        IF NOT _done THEN
            _to_A._sut_A.Invoke();
            _to_A._sut_B.Invoke();
            _to_A();

            IF _to_A._sut_A.Done AND NOT _retBool THEN
                _to_A._sut_A.Abort();
                _to_A._sut_B.Abort();
                _retBool := true;
            END_IF

            _done := _to_A._sut_A.Done AND _to_A._sut_B.Done;
        END_IF

        IF _done THEN
            _to_A._sut_A.ReadOutState();
            _to_A._sut_B.ReadOutState();
            ProbeDoneWhen(_done);
        END_IF
    {endregion}
    {region "T310_TaskError"}
    eTcoTaskTests.TaskError:
        IF NOT _arranged THEN
            IF _plcCycleCounter = 1 THEN
                _to_A.CounterValue_A := _inUint;
                RETURN;
            END_IF

            IF _plcCycleCounter = 2 THEN
                _to_A._sut_A.Invoke();
                RETURN;
            END_IF

            IF _plcCycleCounter > 2 AND _plcCycleCounter <= 5 THEN
                _to_A._sut_A();
                RETURN;
            END_IF

            IF _plcCycleCounter = 6 THEN
                _to_A._sut_A();
                _to_A._sut_A.ReadOutState();
                _arranged := TRUE;
                RETURN;
            END_IF
        END_IF

        IF NOT _done THEN
            IF _plcCycleCounter = 7 THEN
                _to_A.CounterValue_A := _to_A.CounterValue_A + 5;
                _to_A._sut_A();
                _to_A._sut_A.ReadOutState();
            END_IF

            IF _plcCycleCounter > 7 AND _plcCycleCounter <= 7 + _inUint THEN
                _to_A._sut_A();
                _to_A._sut_A.ReadOutState();
            END_IF

            _done := _plcCycleCounter >= 7 + _inUint;
            ProbeDoneWhen(_done);
        END_IF
    {endregion}
    {region "T311_TaskInvokeAfterErrorNoRestoreNoEmptyCycles"}
    eTcoTaskTests.TaskInvokeAfterErrorNoRestoreNoEmptyCycles:
        IF NOT _arranged THEN
            _to_A._sut_A.Invoke();
            _arranged := TRUE;
            RETURN;
        END_IF

        IF NOT _done THEN
            _to_A._sut_A();
            _to_A._sut_A.ReadOutState();
            ProbeDoneWhen(_plcCycleCounter >= 1 + _inUint);
        END_IF
    {endregion}
    {region "T312_TaskInvokeAfterErrorNoRestoreOneEmptyCycle"}
    eTcoTaskTests.TaskInvokeAfterErrorNoRestoreOneEmptyCycle:
        IF NOT _arranged THEN
            IF _plcCycleCounter = 1 THEN
                RETURN;
            END_IF

            IF _plcCycleCounter = 2 THEN
                _to_A._sut_A.Invoke();
                RETURN;
            END_IF
        END_IF

        IF NOT _done THEN
            _to_A._sut_A();
            _to_A._sut_A.ReadOutState();
            _done := _plcCycleCounter >= 2 + _inUint;
            ProbeDoneWhen(_done);
        END_IF
    {endregion}
    {region "T313_TaskInvokeAfterErrorWithRestore"}
    eTcoTaskTests.TaskInvokeAfterErrorWithRestore:
        _to_A._sut_A.Restore();
        _to_A._sut_A.Invoke();
        _to_A._sut_A();
        _to_A._sut_A.ReadOutState();
        _done := TRUE;
        ProbeDoneWhen(_done);
    {endregion}
    {region "T314_TaskAbortDuringExecution"}
    eTcoTaskTests.TaskAbortDuringExecution:
        IF _plcCycleCounter = 1 THEN
            _to_A._sut_A.Restore();
            RETURN;
        END_IF

        IF _plcCycleCounter = 2 THEN
            _to_A._sut_A.Invoke();
            _to_A._sut_A();
            _to_A._sut_A.ReadOutState();
            RETURN;
        END_IF

        IF _plcCycleCounter = 3 THEN
            _to_A._sut_A.Abort();
            _to_A._sut_A();
            _to_A._sut_A.ReadOutState();
            _done := TRUE;
            ProbeDoneWhen(_done);
        END_IF
    {endregion}
    {region "T315_TaskMessage"}
    eTcoTaskTests.TaskMessage:
        _to_A._sut_A.PostMessage(Message := _inString);
        _retString := _to_A._sut_A.GetMessage();
        _done := TRUE;
        ProbeDoneWhen(_done);
    {endregion}
    {region "T316_IdentitiesTest"}
    eTcoTaskTests.IdentitiesTest:
        _runElapsedTimer := TRUE;
        _elapsedTimeETA := UINT_TO_TIME(_inUint);
        _to_A._sut_A.ReadOutIdentities();
        _to_A.ReadOutIdentities();
        ReadOutCycleCounters();
        _done := _elapsedTimeTimer.Q;
        ProbeDoneWhen(_done);
    {endregion}
    {region "T317_CheckAutoRestoreProperties"}
    eTcoTaskTests.CheckAutoRestoreProperties:
        _to_A._tSt_A.ReadOutAutoRestoreProperties();
        _to_A._tSt_B.ReadOutAutoRestoreProperties();
        _to_A._tSt_A._tTt_A.ReadOutAutoRestoreProperties();
        _to_A._tSt_A._tTt_B.ReadOutAutoRestoreProperties();
        _to_A._tSt_B._tTt_A.ReadOutAutoRestoreProperties();
        _to_A._tSt_B._tTt_B.ReadOutAutoRestoreProperties();
        _done := TRUE;
        ProbeDoneWhen(_done);
    {endregion}
    {region "T318_AutoRestoreOnStateChange"}
    eTcoTaskTests.AutoRestoreOnStateChange:
        IF _plcCycleCounter = 1 THEN
            _to_A._tSt_A.ReadOutAutoRestoreProperties();
            _to_A._tSt_B.ReadOutAutoRestoreProperties();
            _to_A._tSt_A._tTt_A.ReadOutAutoRestoreProperties();
            _to_A._tSt_A._tTt_B.ReadOutAutoRestoreProperties();
            _to_A._tSt_B._tTt_A.ReadOutAutoRestoreProperties();
            _to_A._tSt_B._tTt_B.ReadOutAutoRestoreProperties();
            _to_A._tSt_A._tTt_A.ReadOutState();
            _to_A._tSt_B._tTt_B.ReadOutState();
        END_IF

        IF _plcCycleCounter = 2 THEN
            _to_A._tSt_A._tTt_A.Restore();
            _to_A._tSt_B._tTt_B.Restore();
            _to_A._tSt_A._tTt_A.ReadOutState();
            _to_A._tSt_B._tTt_B.ReadOutState();
        END_IF

        IF _plcCycleCounter = 3 THEN
            _to_A._tSt_A._tTt_A.Invoke();
            _to_A._tSt_B._tTt_B.Invoke();
            _to_A._tSt_A._tTt_A();
            _to_A._tSt_B._tTt_B();
            _to_A._tSt_A._tTt_A.ReadOutState();
            _to_A._tSt_B._tTt_B.ReadOutState();
        END_IF

        IF _plcCycleCounter = 4 THEN
            _to_A._tSt_A._tTt_A.Invoke();
            _to_A._tSt_A._tTt_A();
            _to_A._tSt_B._tTt_B();
            _to_A._tSt_A._tTt_A.ReadOutState();
            _to_A._tSt_B._tTt_B.ReadOutState();
        END_IF

        IF _plcCycleCounter = 5 THEN
            _to_A._tSt_A.ChangeState(_to_A._tSt_A._myState);
            _to_A._tSt_B.ChangeState(_to_A._tSt_B._myState);
            _to_A._tSt_A._tTt_A();
            _to_A._tSt_B._tTt_B();
            _to_A._tSt_A._tTt_A.ReadOutState();
            _to_A._tSt_B._tTt_B.ReadOutState();
        END_IF

        _done := _plcCycleCounter = 5;
        ProbeDoneWhen(_done);
    {endregion}
    {region "T320_InvokeDisabledTask"}
    eTcoTaskTests.InvokeDisabledTask:
        IF _plcCycleCounter = 1 THEN
            _to_A._sut_A.Restore();
            _to_A._sut_A.Disable();
            RETURN;
        END_IF

        IF NOT _done THEN
            _to_A._sut_A.Invoke();
            _to_A._sut_A();
            _to_A._sut_A.ReadOutState();
            _done := _plcCycleCounter >= 1 + _inUint;
            ProbeDoneWhen(_done);
        END_IF
    {endregion}
    {region "T321_DisableExecutingTask"}
    eTcoTaskTests.DisableExecutingTask:
        IF _plcCycleCounter = 1 THEN
            _to_A._sut_A.Enable();
            _to_A._sut_A.Invoke();
            _to_A._sut_A();
            _to_A._sut_A.ReadOutState();
            RETURN;
        END_IF

        IF _plcCycleCounter = 2 THEN
            _to_A._sut_A.Disable();
            _to_A._sut_A();
            _to_A._sut_A.ReadOutState();
            RETURN;
        END_IF

        IF _plcCycleCounter = 3 THEN
            _to_A._sut_A.Restore();
            _to_A._sut_A.Enable();
            _to_A._sut_A();
            _to_A._sut_A.ReadOutState();
            RETURN;
        END_IF

        IF _plcCycleCounter = 4 THEN
            _to_A._sut_A.Invoke();
            _to_A._sut_A();
            _to_A._sut_A.ReadOutState();
            RETURN;
        END_IF

        IF _plcCycleCounter = 5 THEN
            _to_A._sut_A.Restore();
            _to_A._sut_A();
            _to_A._sut_A.ReadOutState();
            _done := TRUE;
            ProbeDoneWhen(_done);
        END_IF
    {endregion}
    {region "T322_InvokeTaskThenDisable"}
    eTcoTaskTests.InvokeTaskThenDisable:
        _to_A._sut_A.Invoke();
        _to_A._sut_A.Disable();
        _to_A._sut_A();
        _to_A._sut_A.ReadOutState();
        _done := TRUE;
        ProbeDoneWhen(_done);
    {endregion}
    {region "T323_DisableTaskInErrorStateEnableAndTriggerAgain"}
    eTcoTaskTests.DisableTaskInErrorStateEnableAndTriggerAgain:
        IF _plcCycleCounter = 1 THEN
            _to_A._sut_A.Enable();
            _to_A._sut_A.Invoke();
            _to_A._sut_A();
            _to_A._sut_A.ReadOutState();
            RETURN;
        END_IF

        IF _plcCycleCounter = 2 THEN
            _to_A.CounterValue_A := _to_A.CounterValue_A + 5;
            _to_A._sut_A();
            _to_A._sut_A.ReadOutState();
            RETURN;
        END_IF

        IF _plcCycleCounter = 3 THEN
            _to_A._sut_A.Disable();
            _to_A._sut_A();
            _to_A._sut_A.ReadOutState();
            RETURN;
        END_IF

        IF _plcCycleCounter = 4 THEN
            _to_A._sut_A.Invoke();
            _to_A._sut_A();
            _to_A._sut_A.ReadOutState();
            RETURN;
        END_IF

        IF _plcCycleCounter = 5 THEN
            _to_A._sut_A.Restore();
            _to_A._sut_A.Invoke();
            _to_A._sut_A();
            _to_A._sut_A.ReadOutState();
            _done := TRUE;
            ProbeDoneWhen(_done);
        END_IF
    {endregion}
    {region "T330_ElapsedTypeMeasurement"}
    eTcoTaskTests.ElapsedTypeMeasurement:
        IF _plcCycleCounter = 1 THEN
            _to_A._sut_A.Restore();
            _to_A._sut_A.Enable();
            _to_A._sut_A.Invoke();
            RETURN;
        END_IF

        IF (_to_A._sut_A.Execute()) THEN
            _runElapsedTimer := TRUE;

            IF (_elapsedTimeTimer.Q) THEN
                _to_A._sut_A.DoneWhen(_elapsedTimeTimer.Q);
            END_IF;
        END_IF

        _done := _to_A._sut_A.Done;
        ProbeDoneWhen(_done);
        _elapsedTime := _to_A._sut_A.ElapsedTime;
    {endregion}
    {region "T340_TaskExecutingWithDoneAndErrorStatement"}
    eTcoTaskTests.TaskExecutingWithDoneAndErrorStatement:
        IF _plcCycleCounter = 1 THEN
            _to_A._sut_A.Restore();
            _to_A._sut_A.Enable();
            _to_A._sut_A.Invoke();
            _to_A._sut_A();
            _to_A._sut_A.ReadOutState();
            RETURN;
        END_IF

        _to_A._sut_A();
        _to_A._sut_A.DoneWhen(TRUE);
        _to_A._sut_A.ThrowWhen(TRUE);
        _to_A._sut_A.ReadOutState();
        _done := _to_A._sut_A.Done;
        ProbeDoneWhen(_done);
    {endregion}
    {region "T341_TaskExecutingWithErrorAndDoneStatement"}
    eTcoTaskTests.TaskExecutingWithErrorAndDoneStatement:
        IF _plcCycleCounter = 1 THEN
            _to_A._sut_A.Restore();
            _to_A._sut_A.Enable();
            _to_A._sut_A.Invoke();
            _to_A._sut_A();
            _to_A._sut_A.ReadOutState();
            RETURN;
        END_IF

        _to_A._sut_A();
        _to_A._sut_A.ThrowWhen(TRUE);
        _to_A._sut_A.DoneWhen(TRUE);
        _to_A._sut_A.ReadOutState();
        _done := _to_A._sut_A.Done;
        ProbeDoneWhen(_done);			 
{endregion}
	 eTcoTaskTests.TaskExecuteMethodNotCalled:
	 	_to_A._sut_A.Invoke().Done;
	eTcoTaskTests.TaskExecuteMethodCalled :
		_to_A._sut_A.Invoke().Done;
		_to_A._sut_A.Execute();
END_CASE
END_METHOD

METHOD INTERNAL ReadOutCycleCounters
_startCycles		:=		THIS^.StartCycleCount;
_endCycles			:=		THIS^.EndCycleCount;

_myIdentity			:= 		THIS^.Identity;
END_METHOD

END_FUNCTION_BLOCK

// ---- Tests/TcoTask/PlcExecuted/TcoTaskPlcTestObject.TcPOU
FUNCTION_BLOCK TcoTaskPlcTestObject EXTENDS TcoCore.TcoObject
VAR
	_myIdentity				:	ULINT;
	_myContextIdentity		:	ULINT;
	_myContextStartCount 	:	ULINT;
	_myContextEndCount		:	ULINT;
	_myParentIdentity		:	ULINT;
    _sut_A : TcoTaskPlcTest(THIS^);
    _sut_B : TcoTaskPlcTest(THIS^);
	_tSt_A:TcoTaskPlcTestState(THIS^, eRestoreMode.AutoRestoreMembers);
	_tSt_B:TcoTaskPlcTestState(THIS^, eRestoreMode.None);
END_VAR

_sut_A();
_sut_B();

PROPERTY CounterValue_A : ULINT
GET
CounterValue_A := _sut_A.CounterValue;
END_GET
SET
_sut_A.CounterValue := CounterValue_A;
END_SET
END_PROPERTY

PROPERTY CounterValue_B : ULINT
GET
CounterValue_B := _sut_B.CounterValue;
END_GET
SET
_sut_B.CounterValue := CounterValue_B;
END_SET
END_PROPERTY

{attribute 'TcRpcEnable'}
METHOD INTERNAL ReadOutIdentities
_myIdentity			:=	THIS^.Identity;

_myContextIdentity	:=	THIS^.Context.Identity;
		
_myContextStartCount :=	THIS^.Context.StartCycleCount;

_myContextEndCount	:=	THIS^.Context.EndCycleCount;

_myParentIdentity	:=	THIS^.Parent.Identity;
END_METHOD

END_FUNCTION_BLOCK

// ---- Tests/TcoTask/PlcExecuted/TcoTaskPlcTest.TcPOU
FUNCTION_BLOCK TcoTaskPlcTest EXTENDS TcoCore.TcoTask
VAR
    _isBusy : BOOL;
    _isError : BOOL;
    _isDone : BOOL;
    _isReady : BOOL;
    _isInvokeRequestTrue : BOOL;
    _counterSetValue : ULINT;
    _counterValue : ULINT;
    _invokeCounter : ULINT;
    _executeCounter : ULINT;
    _doneCounter : ULINT;
    _invokeRisingEdgeCounter : ULINT;
    _executeRisingEdgeCounter : ULINT;
    _doneRisingEdgeCounter : ULINT;
    _previousState : eTaskState;
    _counterValuePV : ULINT;
    _myIdentity : ULINT;
    _myContextIdentity : ULINT;
    _myContextStartCount : ULINT;
    _myContextEndCount : ULINT;
    _myParentIdentity : ULINT;
    _autoRestoreByMyParentEnabled : BOOL;
    _onErrorCounter : ULINT;
    _whileErrorCounter : ULINT;
    _onStartCounter : ULINT;
END_VAR

IF(THIS^._taskState = eTaskState.Requested) THEN
	_invokeCounter := _invokeCounter + 1; 
END_IF;

IF(THIS^._taskState = eTaskState.Requested AND _PreviousState <> eTaskState.Requested) THEN
	_counterValue	:=	_counterSetValue;
	_counterValuePV := _counterValue;
	_invokeRisingEdgeCounter := _invokeRisingEdgeCounter + 1;
END_IF

IF(THIS^._taskState = eTaskState.Busy AND _previousState <> eTaskState.Busy) THEN
	_executeRisingEdgeCounter := _executeRisingEdgeCounter + 1;
END_IF

_previousState	:=	THIS^._taskState;

IF(Execute()) THEN
	_executeCounter := _executeCounter + 1;	
	_counterValue := _counterValue - 1;
	DoneWhen(_counterValue <= 0);			
	ThrowWhen(ABS(_counterValuePV -_counterValue) > 1);
	_CounterValuePV := _counterValue;
END_IF

IF(THIS^._taskState = eTaskState.Done) THEN
	_doneCounter := _doneCounter + 1; 
END_IF;

IF(THIS^._taskState = eTaskState.Done AND _previousState <> eTaskState.Done) THEN
	_doneRisingEdgeCounter := _doneRisingEdgeCounter + 1; 
END_IF

PROPERTY CounterValue : ULINT
GET
CounterValue := _counterValue;
END_GET
SET
_counterValue := CounterValue;
END_SET
END_PROPERTY

METHOD INTERNAL Disable
THIS^.Enabled := FALSE;
END_METHOD

METHOD INTERNAL Enable
THIS^.Enabled := TRUE;
END_METHOD

METHOD INTERNAL GetMessage : STRING
GetMessage := SUPER^._messenger._mime.Text;
END_METHOD

METHOD PROTECTED OnError
_onErrorCounter := _onErrorCounter +1;
END_METHOD

METHOD PROTECTED OnStart
_onStartCounter := _onStartCounter +1;
END_METHOD

METHOD INTERNAL PostMessage
VAR_INPUT
	Message	:	STRING;
END_VAR
THIS^.Messenger.Post(Message ,eMessageCategory.Error);
END_METHOD

{attribute 'TcRpcEnable'}
METHOD INTERNAL ReadOutAutoRestoreProperties
_autoRestoreByMyParentEnabled	:= THIS^.AutoRestorable;
END_METHOD

{attribute 'TcRpcEnable'}
METHOD INTERNAL ReadOutIdentities
_myIdentity			:=	THIS^.Identity;
 
_myContextIdentity	:=	THIS^.Context.Identity;
		
_myContextStartCount :=	THIS^.Context.StartCycleCount;
 
_myContextEndCount	:=	THIS^.Context.EndCycleCount;
 
_myParentIdentity	:=	THIS^.Parent.Identity;
END_METHOD

{attribute 'TcRpcEnable'}
METHOD INTERNAL ReadOutState
_isBusy					:=	THIS^.Busy;	
_isError				:=	THIS^.Error;	
_isDone					:=	THIS^.Done;	
_isReady				:=	THIS^.Ready;
_isInvokeRequestTrue 	:=	THIS^._invokeRequest;
END_METHOD

{attribute 'TcRpcEnable'}
METHOD INTERNAL SetInvokeRequest
THIS^._invokeRequest := TRUE;
END_METHOD

{attribute 'TcRpcEnable'}
METHOD INTERNAL SetPreviousStateToReady
THIS^._previousState := eTaskState.Ready;
END_METHOD

(*~
	<docu>
		<summary>
			Executes until task is in ```Error``` state .
		</summary>			
	</docu>	
~*)
METHOD PROTECTED WhileError
_whileErrorCounter := _whileErrorCounter + 1;
END_METHOD

END_FUNCTION_BLOCK

// ---- Tests/TcoTask/PlcExecuted/TcoTaskPlcTestState.TcPOU
FUNCTION_BLOCK TcoTaskPlcTestState EXTENDS TcoState
VAR
    _myIdentity : ULINT;
    _myContextIdentity : ULINT;
    _myContextStartCount : ULINT;
    _myContextEndCount : ULINT;
    _myParentIdentity : ULINT;
    _myState : INT;
    _tTt_A : TcoTaskPlcTest(THIS^);
    _tTt_B : TcoTaskPlcTest(THIS^);
    _onStateChangeCounter : INT;
    _autoRestoreToMyChildsEnabled : BOOL;
    _autoRestoreByMyParentEnabled : BOOL;
END_VAR

METHOD PROTECTED OnStateChange 
VAR_INPUT
	PreviousState	: INT;
	NewState 		: INT;
END_VAR
VAR
	message	:	STRING;
END_VAR
_onStateChangeCounter	:=	_onStateChangeCounter + 1;

message := CONCAT('My state has been change from ', INT_TO_STRING(PreviousState));
message := CONCAT(message, ' to the new state ');
message := CONCAT(message, INT_TO_STRING(NewState));
message := CONCAT(message, '.');

THIS^.Messenger.Post(message,eMessageCategory.Debug);

SUPER^.OnStateChange(PreviousState,NewState);
END_METHOD

{attribute 'TcRpcEnable'}
METHOD INTERNAL ReadOutAutoRestoreProperties
_autoRestoreToMyChildsEnabled	:= THIS^.IsAutoRestoreEnabled;
_autoRestoreByMyParentEnabled	:= THIS^.AutoRestorable;
END_METHOD

{attribute 'TcRpcEnable'}
METHOD INTERNAL ReadOutIdentities
_myIdentity			:=	THIS^.Identity;

_myContextIdentity	:=	THIS^.Context.Identity;

_myParentIdentity	:=	THIS^.Parent.Identity;
		
_myContextStartCount :=	THIS^.Context.StartCycleCount;

_myContextEndCount	:=	THIS^.Context.EndCycleCount;
END_METHOD

{attribute 'TcRpcEnable'}
METHOD INTERNAL ReadOutState
_myState			:=	THIS^.State;

THIS^._tTt_A.ReadOutState();
THIS^._tTt_B.ReadOutState();
END_METHOD

{attribute 'TcRpcEnable'}
METHOD INTERNAL TriggerChangeState
VAR_INPUT
	NewState : INT;
END_VAR
THIS^.ChangeState(NewState);
END_METHOD

{attribute 'TcRpcEnable'}
METHOD INTERNAL TriggerChangeStateWithObjectRestore
VAR_INPUT
	NewState : INT;
END_VAR
THIS^.ChangeState(NewState).RestoreObject(THIS^._tTt_A).RestoreObject(THIS^._tTt_B);
END_METHOD

{attribute 'TcRpcEnable'}
METHOD INTERNAL TriggerRestore
THIS^.Restore();
END_METHOD

{attribute 'TcRpcEnable'}
METHOD INTERNAL TriggerTaskInvoke
THIS^._tTt_A.Invoke();

THIS^._tTt_B.Invoke();
END_METHOD

END_FUNCTION_BLOCK

// ---- Tests/TcoToggleTask/TcoToggleTaskTestContext.TcPOU
FUNCTION_BLOCK TcoToggleTaskTestContext EXTENDS TcoCore._internals_TcoContext
VAR
    _sut 		:	TcoToggleTaskTests(THIS^, TRUE);
	_bool		:	BOOL;
	_string		:	STRING;
	_done		:	BOOL;
END_VAR

METHOD PROTECTED Main
CASE _testId OF
	eTcoToggleTaskTests.Reinit:
		_sut.FB_init(TRUE, FALSE, THIS^,_bool);
		_done := TRUE;
		
	eTcoToggleTaskTests.CleanUp:
		IF NOT _done THEN
			_sut._messenger.Clear();
			_done := TRUE;
		END_IF
		
	eTcoToggleTaskTests.Message:
		IF NOT _done THEN
			_sut.Messenger.Error(_string);
			_done := TRUE;
		END_IF
		
	eTcoToggleTaskTests.TriggerToggleWhileRunNotCalled:
		IF NOT _done THEN
			_sut._messenger.Clear();
			_sut.Toggle();
			_done := TRUE;	
		END_IF

	eTcoToggleTaskTests.TriggerToggleWhileDisabled:
		IF NOT _done THEN
			_sut.Run();
			_sut._messenger.Clear();
			_sut.Enabled := FALSE;
			_sut.Toggle();
			_done := TRUE;	
		END_IF

	eTcoToggleTaskTests.TriggerToggleWhileEnabled:
		IF NOT _done THEN
			_sut.Run();
			_sut._messenger.Clear();
			_sut.Enabled := TRUE;
			_sut.Toggle();
			_done := TRUE;	
		END_IF

	eTcoToggleTaskTests.TriggerOnWhileRunNotCalled:
		IF NOT _done THEN
			_sut._messenger.Clear();
			_sut.On();
			_done := TRUE;	
		END_IF

	eTcoToggleTaskTests.TriggerOnWhileDisabled:
		IF NOT _done THEN
			_sut.Run();
			_sut._messenger.Clear();
			_sut.Enabled := FALSE;
			_sut.On();
			_done := TRUE;	
		END_IF

	eTcoToggleTaskTests.TriggerOnWhileEnabled:
		IF NOT _done THEN
			_sut.Run();
			_sut._messenger.Clear();
			_sut.Enabled := TRUE;
			_sut.On();
			_done := TRUE;	
		END_IF

	eTcoToggleTaskTests.TriggerOffWhileRunNotCalled:
		IF NOT _done THEN
			_sut._messenger.Clear();
			_sut.Toggle();
			_done := TRUE;	
		END_IF

	eTcoToggleTaskTests.TriggerOffWhileDisabled:
		IF NOT _done THEN
			_sut.Run();
			_sut._messenger.Clear();
			_sut.Enabled := FALSE;
			_sut.Off();
			_done := TRUE;	
		END_IF

	eTcoToggleTaskTests.TriggerOffWhileEnabled:
		IF NOT _done THEN
			_sut.Run();
			_sut._messenger.Clear();
			_sut.Enabled := TRUE;
			_sut.Off();
			_done := TRUE;	
		END_IF

		
END_CASE
END_METHOD

END_FUNCTION_BLOCK

// ---- Tests/TcoToggleTask/TcoToggleTaskTests.TcPOU
FUNCTION_BLOCK TcoToggleTaskTests EXTENDS TcoCore.TcoToggleTask
VAR
	_isOn							:	BOOL;	
	_isOff							:	BOOL;	
	_isEnabled						:	BOOL;	
	_isToggleRequestTrue			:	BOOL;		
	_counterValue					:	ULINT;
	_counterValuePV					:	ULINT;
	_toggleCounter					:	ULINT;
	_runCounter						:	ULINT;
	_onFtrigCounter					:	ULINT;	
	_onRtrigCounter					:	ULINT;	
	_onCounter						:	ULINT;
	_offCounter						:	ULINT;
	_onStateChangeCounter			:	ULINT;
	_taskOnCounter					:	ULINT;
	_taskOffCounter					:	ULINT;
	_stateChangedCounter			:	ULINT;

	_previousState					:	BOOL;
	_myIdentity						:	ULINT;
	_myContextIdentity				:	ULINT;
	_myContextStartCount 			:	ULINT;
	_myContextEndCount				:	ULINT;	
	_myParentIdentity				:	ULINT;
END_VAR

ExecutionBody();

METHOD INTERNAL Disable
THIS^.Enabled := FALSE;
END_METHOD

METHOD INTERNAL Enable
THIS^.Enabled := TRUE;
END_METHOD

{attribute 'TcRpcEnable'}
METHOD INTERNAL ExecutionBody
Run();

_runCounter := _runCounter + 1;	

IF _previousState <> THIS^.State THEN
	_stateChangedCounter := _stateChangedCounter + 1;
END_IF; 
_previousState	:=	THIS^.State;
END_METHOD

{attribute 'TcRpcEnable'}
METHOD INTERNAL GetMessage : STRING
GetMessage := SUPER^._messenger._mime.Text;
END_METHOD

METHOD PROTECTED Main
VAR
	
END_VAR
END_METHOD

(*~
	<docu>
		<summary>
			Executes when toggle task changes its state from '''TRUE''' to '''FALSE'''.
		</summary>			
	</docu>	
~*)
METHOD PROTECTED OnFtrig
_onFtrigCounter := _onFtrigCounter + 1;
END_METHOD

(*~
	<docu>
		<summary>
			Executes when toggle task changes its state from '''FALSE''' to '''TRUE'''.
		</summary>			
	</docu>	
~*)
METHOD PROTECTED OnRtrig
_onRtrigCounter := _onRtrigCounter + 1;
END_METHOD

(*~
	<docu>
		<summary>
			Executes when toggle task changes its state .
		</summary>			
	</docu>	
~*)
METHOD PROTECTED OnStateChange
_onStateChangeCounter := _onStateChangeCounter + 1;
END_METHOD

{attribute 'TcRpcEnable'}
METHOD INTERNAL PostMessage
VAR_INPUT
	Message	:	STRING;
END_VAR
THIS^.Messenger.Post(Message ,eMessageCategory.Error);
END_METHOD

{attribute 'TcRpcEnable'}
METHOD INTERNAL ReadOutIdentities
_myIdentity			:=	THIS^.Identity;
 
_myContextIdentity	:=	THIS^.Context.Identity;
		
_myContextStartCount :=	THIS^.Context.StartCycleCount;
 
_myContextEndCount	:=	THIS^.Context.EndCycleCount;
 
_myParentIdentity	:=	THIS^.Parent.Identity;
END_METHOD

{attribute 'TcRpcEnable'}
METHOD INTERNAL ReadOutState
_isOn				    :=	THIS^.IsOn;	
_isOff				   	:=	THIS^.IsOff;	
_isEnabled				:=	THIS^.Enabled;
_isToggleRequestTrue	:=	THIS^._toggleRequest;
END_METHOD

{attribute 'TcRpcEnable'}
METHOD INTERNAL SetPreviousState
VAR_INPUT
	inValue : BOOL;
END_VAR
THIS^._previousState := inValue;
END_METHOD

{attribute 'TcRpcEnable'}
METHOD INTERNAL SetState
VAR_INPUT
	inState	:	BOOL;
END_VAR
THIS^._state := inState;
END_METHOD

{attribute 'TcRpcEnable'}
METHOD INTERNAL SetToggleRequest
THIS^._toggleRequest := TRUE;
END_METHOD

(*~
	<docu>
		<summary>
			Executes when toggle task is in ```Off``` state .
		</summary>			
	</docu>	
~*)
METHOD PROTECTED TaskOff
_taskOffCounter := _taskOffCounter + 1;

_counterValue := _counterValue - 1;
_CounterValuePV := _counterValue;
END_METHOD

(*~
	<docu>
		<summary>
			Executes when toggle task is in  ```On``` state .
		</summary>			
	</docu>	
~*)
METHOD PROTECTED TaskOn
_taskOnCounter := _taskOnCounter + 1;

_counterValue := _counterValue + 1;
_CounterValuePV := _counterValue;
END_METHOD

{attribute 'TcRpcEnable'}
METHOD INTERNAL TriggerOff
THIS^.Off();
_offCounter := _offCounter + 1;
END_METHOD

{attribute 'TcRpcEnable'}
METHOD INTERNAL TriggerOn
THIS^.On();
_onCounter := _onCounter + 1;
END_METHOD

{attribute 'TcRpcEnable'}
METHOD INTERNAL TriggerToggle
THIS^.Toggle();
_toggleCounter := _toggleCounter + 1;
END_METHOD

END_FUNCTION_BLOCK

// ---- Tests/TcoComponent/PlcExecuted/TcoComponentTestContext.TcPOU
FUNCTION_BLOCK TcoComponentTestContext EXTENDS TcoCore._internals_TcoContext
VAR	
    _sut : TestComponent(THIS^);
	{attribute addProperty Name "--Some IO signal"}
	_signal : BOOL;	
END_VAR

METHOD PROTECTED Main
CASE _testId OF
	eTcoComponentTests.GetSignalInfo:
		_sut(_signal := _signal);
END_CASE
END_METHOD

END_FUNCTION_BLOCK

// ---- Tests/TcoComponent/PlcExecuted/TestComponent.TcPOU
FUNCTION_BLOCK TestComponent EXTENDS TcoCore.TcoComponent
VAR_IN_OUT
	_signal : BOOL;
END_VAR
VAR
	_signalInfo : TcoCore.TcoSignalInfo;
END_VAR

_signalInfo.GetSignalInfo(SIZEOF(_signal), ADR(_signal));

(*~
	<docu>
		<summary>
			Restores this instance to the Ready state. Can be called explicitly or from within one of the restore mechanisms.	
		</summary>			
	</docu>	
~*)
METHOD  Restore : ITcoRestorable
END_METHOD

(*~
	<docu>
		<summary>
		    Custom service (manual, maintenance) logic.
			This method must be implemented in derived class.
		</summary>			
	</docu>	
~*)
METHOD PROTECTED  ServiceMode
END_METHOD

END_FUNCTION_BLOCK

// ---- Tests/TcoRemoteTask/PlcExecuted/TcoRemoteTaskTestContext.TcPOU
FUNCTION_BLOCK TcoRemoteTaskTestContext EXTENDS TcoCore._internals_TcoContext
VAR
	_sut : TcoRemoteTaskTest(THIS^);
    _invokeInitializedCSharpMethodDone : BOOL;
    _invokeNotInitializedCSharpMethodDone : BOOL;
    _exceptionInMethodWillResultInExceptionDone : BOOL;
	_sharedVariable : INT;
	
END_VAR

METHOD PROTECTED Main

CASE _testId OF
    0:
        _invokeInitializedCSharpMethodDone := FALSE;
        _invokeNotInitializedCSharpMethodDone := FALSE;
        _exceptionInMethodWillResultInExceptionDone := FALSE;
    eTcoRemoteTaskTests.RestoreTasks:
        _sut._invokeInitializedCSharpMethod.Restore();
        _sut._invokeNotInitializedCSharpMethod.Restore();
        _sut._exceptionInMethodWillResultInException.Restore();
    eTcoRemoteTaskTests.InvokeInitializedCSharpMethod:
        _invokeInitializedCSharpMethodDone := _sut._invokeInitializedCSharpMethod.Invoke().Done;
    eTcoRemoteTaskTests.InvokeNotInitializedCSharpMethod:
        _invokeNotInitializedCSharpMethodDone := _sut._invokeNotInitializedCSharpMethod.Invoke().Error;
    eTcoRemoteTaskTests.ExceptionInMethodWillResultInException:
        _exceptionInMethodWillResultInExceptionDone := _sut._exceptionInMethodWillResultInException.Invoke().Error;
END_CASE

_sut();
END_METHOD

END_FUNCTION_BLOCK

// ---- Tests/TcoRemoteTask/PlcExecuted/TcoRemoteTaskTest.TcPOU
FUNCTION_BLOCK TcoRemoteTaskTest EXTENDS TcoCore.TcoObject
VAR
	_invokeInitializedCSharpMethod : TcoCore.TcoRemoteTask(THIS^);
    _invokeNotInitializedCSharpMethod : TcoCore.TcoRemoteTask(THIS^);
    _exceptionInMethodWillResultInException : TcoCore.TcoRemoteTask(THIS^);
END_VAR

_invokeInitializedCSharpMethod();
_invokeNotInitializedCSharpMethod();
_exceptionInMethodWillResultInException();

END_FUNCTION_BLOCK

// ---- Tests/TcoSequencer/PlcExecuted/TcoSequencerTestContext.TcPOU
FUNCTION_BLOCK TcoSequencerTestContext EXTENDS TcoCore._internals_TcoContext
VAR
    _sut_A : TcoSequencerTestType(THIS^, eRestoreMode.AutoRestoreMembers);
    _sut_N : TcoSequencerTestType(THIS^, eRestoreMode.None);

    _elapsedTimeETA : TIME;
    _elapsedTime : TIME;
    _runElapsedTimer : BOOL;
    _elapsedTimeTimer : Tc2_Standard.TON;

	_runOneStep							:	BOOL;
	_runAllSteps						:	BOOL;
	_finishStep							:	BOOL;
	_stepId								:	INT;
	_enabled							:	BOOL;
	_stepDescription					:	STRING(254);	
	_currentStepId						:	INT;
	_currentStepDescription				:	STRING(254);
    _totalStepNumber : UINT;
	_reqStep : INT;
    _reqStepNotExists : INT;

    _done : BOOL;
    _arranged : BOOL;
	_startCycles			:	ULINT;
	_endCycles				:	ULINT;	
	_myIdentity				:	ULINT;	
	_initReqStepCycle		:	UINT;
	_cycles					:	UINT;
	_cyclicCycles :	UINT;
    _stepInEvents :	UINT;

END_VAR

{attribute 'TcRpcEnable'}
METHOD _ClearPlcCycleCounter
ClearPlcCycleCounter();
END_METHOD

METHOD PROTECTED Main
VAR
	i:INT;
END_VAR
_elapsedTimeTimer(IN := _runElapsedTimer, PT := _elapsedTimeETA);

CASE _testId OF
    {region "CallSequencerBodiesOnly"}
    eTcoSequencerTests.CallSequencerBodiesOnly:
        _sut_A.TcoSequencerTest := eTcoSequencerTests.CallSequencerBodiesOnly;
        _sut_N.TcoSequencerTest := eTcoSequencerTests.CallSequencerBodiesOnly;
        _sut_A.Run();
        _sut_N.Run();
    {endregion}
    {region "RestoreSequencers"}
    eTcoSequencerTests.RestoreSequencers:
        IF NOT _arranged THEN
            _sut_A.Restore();
            _sut_N.Restore();
            _arranged := _sut_A._restoringSequence AND _sut_N._restoringSequence;
        END_IF

        IF _arranged AND NOT _done THEN
            _sut_A.TcoSequencerTest := eTcoSequencerTests.RestoreSequencers;
            _sut_N.TcoSequencerTest := eTcoSequencerTests.RestoreSequencers;
            _sut_A.Run();
            _sut_N.Run();

            _done :=
                NOT _sut_A._restoringSequence AND NOT _sut_N._restoringSequence AND NOT _sut_A._sequencerHasError AND NOT _sut_N._sequencerHasError;
        END_IF

        ProbeDoneWhen(_done);
    {endregion}
    {region "T500_NumberOfStepsCount"}
    eTcoSequencerTests.NumberOfStepsCount:
        IF NOT _arranged THEN
            _sut_A.SetCyclicMode(); //Set sequencer into the cyclic mode
            _sut_N.SetCyclicMode(); //Set sequencer into the cyclic mode
            _sut_A.SetSequenceAsChecked(); //Set sequence as checked, so no StepID uniqueness is performed on next sequence execution
            _sut_N.SetSequenceAsChecked(); //Set sequence as checked, so no StepID uniqueness is performed on next sequence execution
            _sut_A.ClearNumberOfSteps(); //Clear internal flow step counters, so number of steps is going to be counted again on next sequence run
            _sut_N.ClearNumberOfSteps(); //Clear internal flow step counters, so number of steps is going to be counted again on next sequence run

            _sut_A.SetCurrentStep(_currentStepId,
                _currentStepDescription); //Set the StepId so as the StepDescription to the current step of the sequencer

            _sut_N.SetCurrentStep(_currentStepId,
                _currentStepDescription); //Set the StepId so as the StepDescription to the current step of the sequencer

            _sut_A.SaveNumberOfStepsInSequence();
            _sut_N.SaveNumberOfStepsInSequence();
            _sut_A.TcoSequencerTest := eTcoSequencerTests.NumberOfStepsCount;
            _sut_N.TcoSequencerTest := eTcoSequencerTests.NumberOfStepsCount;
            _sut_A.TotalStepNumber := _totalStepNumber;
            _sut_N.TotalStepNumber := _totalStepNumber;
            _sut_A.FinishStep := FALSE;
            _sut_N.FinishStep := FALSE;
            _arranged := TRUE;
            RETURN;
        END_IF

        IF NOT _done THEN
            _sut_A.Run();
            _sut_N.Run();
            _sut_A.SaveNumberOfStepsInSequence();
            _sut_N.SaveNumberOfStepsInSequence();
            _done := TRUE;
        END_IF

        IF _done THEN
            ProbeDoneWhen(_done);
        END_IF
    {endregion}
    {region "T501_ExecutionInOnePLCcycle"}
    eTcoSequencerTests.ExecutionInOnePLCcycle:
        _sut_A.TcoSequencerTest := eTcoSequencerTests.ExecutionInOnePLCcycle;
        _sut_N.TcoSequencerTest := eTcoSequencerTests.ExecutionInOnePLCcycle;
        _sut_A.SetCyclicMode(); //Set sequencer into the cyclic mode
        _sut_N.SetCyclicMode(); //Set sequencer into the cyclic mode
        _sut_A.TotalStepNumber := _totalStepNumber;
        _sut_N.TotalStepNumber := _totalStepNumber;
        _sut_A.Run();
        _sut_N.Run();
        _done := TRUE;
        ProbeDoneWhen(_done);
    {endregion}
    {region "T502_OnStepCompleted"}
    eTcoSequencerTests.OnStepCompleted:
        _sut_A.TcoSequencerTest := eTcoSequencerTests.OnStepCompleted;
        _sut_N.TcoSequencerTest := eTcoSequencerTests.OnStepCompleted;
        _sut_A.TotalStepNumber := _totalStepNumber;
        _sut_N.TotalStepNumber := _totalStepNumber;
        _sut_A.Run();
        _sut_N.Run();
        _sut_A.SaveNumberOfStepsInSequence();
        _sut_N.SaveNumberOfStepsInSequence();
        _done := TRUE;
        ProbeDoneWhen(_done);
    {endregion}
    {region "T503_OnSequenceCompleted"}
    eTcoSequencerTests.OnSequenceCompleted:
        _sut_A.TcoSequencerTest := eTcoSequencerTests.OnSequenceCompleted;
        _sut_N.TcoSequencerTest := eTcoSequencerTests.OnSequenceCompleted;
        _sut_A.TotalStepNumber := _totalStepNumber;
        _sut_N.TotalStepNumber := _totalStepNumber;
        _sut_A.Run();
        _sut_N.Run();
        _done := TRUE;
        ProbeDoneWhen(_done);
    {endregion}
    {region "T504_RestoreChildBetweenSteps"}
    eTcoSequencerTests.RestoreChildBetweenSteps:
        IF NOT _arranged THEN
            _sut_A.TcoSequencerTest := eTcoSequencerTests.RestoreChildBetweenSteps;
            _sut_N.TcoSequencerTest := eTcoSequencerTests.RestoreChildBetweenSteps;
            _sut_A.TotalStepNumber := _totalStepNumber;
            _sut_N.TotalStepNumber := _totalStepNumber;
            _arranged := TRUE;
            RETURN;
        END_IF;

        _sut_A.Run();
        _sut_N.Run();
        _done := TRUE;
        ProbeDoneWhen(_done);
    {endregion}
    {region "T505_OnStateChangeWithRestoreCallInside"}
    eTcoSequencerTests.OnStateChangeWithRestoreCallInside:
        IF NOT _arranged THEN
            _sut_A.SetCyclicMode(); //Set sequencer into the cyclic mode
            _sut_N.SetCyclicMode(); //Set sequencer into the cyclic mode
            _sut_A.SetSequenceAsChecked(); //Set sequence as checked, so no StepID uniqueness is performed on next sequence execution
            _sut_N.SetSequenceAsChecked(); //Set sequence as checked, so no StepID uniqueness is performed on next sequence execution
            _sut_A.SetNumberOfSteps(_totalStepNumber); //Set numberOfSteps to the testing instance
            _sut_N.SetNumberOfSteps(_totalStepNumber); //Set numberOfSteps to the testing instance
            _sut_A.TcoSequencerTest := eTcoSequencerTests.OnStateChangeWithRestoreCallInside;
            _sut_N.TcoSequencerTest := eTcoSequencerTests.OnStateChangeWithRestoreCallInside;
            _sut_A.TotalStepNumber := _totalStepNumber;
            _sut_N.TotalStepNumber := _totalStepNumber;
            _sut_A.FinishStep := FALSE;
            _sut_N.FinishStep := FALSE;
            _plcCycleCounter := 0;
            _arranged := TRUE;
            RETURN;
        END_IF

        IF NOT _done THEN
            IF _plcCycleCounter = 1 THEN
                _sut_A.CallRestoreInOnStateChange := FALSE;
                _sut_N.CallRestoreInOnStateChange := FALSE;
            ELSE
                _sut_A.CallRestoreInOnStateChange := TRUE;
                _sut_N.CallRestoreInOnStateChange := TRUE;
                _sut_A.FinishStep := TRUE;
                _sut_N.FinishStep := TRUE;
            END_IF

            _sut_A.Run();
            _sut_N.Run();
        END_IF

        _done := _plcCycleCounter >= 2;

        IF _done THEN
            _sut_A.CallRestoreInOnStateChange := FALSE;
            _sut_N.CallRestoreInOnStateChange := FALSE;
            ProbeDoneWhen(_done);
        END_IF
    {endregion}
    {region "T506_MinStepId"}
    eTcoSequencerTests.MinStepId:
        IF NOT _arranged THEN
            _sut_A.SetCyclicMode(); //Set sequencer into the cyclic mode
            _sut_N.SetCyclicMode(); //Set sequencer into the cyclic mode
            _sut_A.SetSequenceAsChecked(); //Set sequence as checked, so no StepID uniqueness is performed on next sequence execution
            _sut_N.SetSequenceAsChecked(); //Set sequence as checked, so no StepID uniqueness is performed on next sequence execution
            _sut_A.SetNumberOfSteps(_totalStepNumber); //Set numberOfSteps to the testing instance
            _sut_N.SetNumberOfSteps(_totalStepNumber); //Set numberOfSteps to the testing instance
            _sut_A.TcoSequencerTest := eTcoSequencerTests.MinStepId;
            _sut_N.TcoSequencerTest := eTcoSequencerTests.MinStepId;
            _sut_A.TotalStepNumber := _totalStepNumber;
            _sut_N.TotalStepNumber := _totalStepNumber;
            _sut_A.FinishStep := FALSE;
            _sut_N.FinishStep := FALSE;
            _plcCycleCounter := 0;
            _arranged := TRUE;
            RETURN;
        END_IF

        IF NOT _done THEN
            _sut_A.StepId := _currentStepId;
            _sut_N.StepId := _currentStepId;
            _sut_A.Run();
            _sut_N.Run();
        END_IF

        _done := TRUE;
        ProbeDoneWhen(_done);
    {endregion}
    {region "T507_MaxStepId"}
    eTcoSequencerTests.MaxStepId:
        IF NOT _arranged THEN
            _sut_A.SetCyclicMode(); //Set sequencer into the cyclic mode
            _sut_N.SetCyclicMode(); //Set sequencer into the cyclic mode
            _sut_A.SetSequenceAsChecked(); //Set sequence as checked, so no StepID uniqueness is performed on next sequence execution
            _sut_N.SetSequenceAsChecked(); //Set sequence as checked, so no StepID uniqueness is performed on next sequence execution
            _sut_A.SetNumberOfSteps(_totalStepNumber); //Set numberOfSteps to the testing instance
            _sut_N.SetNumberOfSteps(_totalStepNumber); //Set numberOfSteps to the testing instance
            _sut_A.TcoSequencerTest := eTcoSequencerTests.MaxStepId;
            _sut_N.TcoSequencerTest := eTcoSequencerTests.MaxStepId;
            _sut_A.TotalStepNumber := _totalStepNumber;
            _sut_N.TotalStepNumber := _totalStepNumber;
            _sut_A.FinishStep := FALSE;
            _sut_N.FinishStep := FALSE;
            _plcCycleCounter := 0;
            _arranged := TRUE;
            RETURN;
        END_IF

        IF NOT _done THEN
            _sut_A.StepId := _currentStepId;
            _sut_N.StepId := _currentStepId;
            _sut_A.Run();
            _sut_N.Run();
        END_IF

        _done := TRUE;
        ProbeDoneWhen(_done);
    {endregion}
    {region "T508_RequestStepToFirstStepWithStepId0"}
    eTcoSequencerTests.RequestStepToFirstStepWithStepId0:
        IF NOT _arranged THEN
            _sut_A.SetCyclicMode(); //Set sequencer into the cyclic mode
            _sut_N.SetCyclicMode(); //Set sequencer into the cyclic mode
            _sut_A.SetSequenceAsChecked(); //Set sequence as checked, so no StepID uniqueness is performed on next sequence execution
            _sut_N.SetSequenceAsChecked(); //Set sequence as checked, so no StepID uniqueness is performed on next sequence execution
            _sut_A.SetNumberOfSteps(_totalStepNumber); //Set numberOfSteps to the testing instance
            _sut_N.SetNumberOfSteps(_totalStepNumber); //Set numberOfSteps to the testing instance
            _sut_A.TcoSequencerTest := eTcoSequencerTests.RequestStepToFirstStepWithStepId0;
            _sut_N.TcoSequencerTest := eTcoSequencerTests.RequestStepToFirstStepWithStepId0;
            _sut_A.TotalStepNumber := _totalStepNumber;
            _sut_N.TotalStepNumber := _totalStepNumber;
            _sut_A.FinishStep := TRUE;
            _sut_N.FinishStep := TRUE;
            _plcCycleCounter := 0;
            _arranged := TRUE;
            RETURN;
        END_IF

        IF NOT _done THEN
            IF _plcCycleCounter > 1 THEN
                _sut_A.FinishStep := FALSE;
                _sut_N.FinishStep := FalsE;
            END_IF

            _sut_A.Run();
            _sut_N.Run();
        END_IF

        _done := _plcCycleCounter > 1;
        ProbeDoneWhen(_done);
    {endregion}
    {region "T509_RequestStep"}
    eTcoSequencerTests.RequestStep:
        IF NOT _arranged THEN
            _sut_A.SetCyclicMode(); //Set sequencer into the cyclic mode
            _sut_N.SetCyclicMode(); //Set sequencer into the cyclic mode
            _sut_A.SetSequenceAsChecked(); //Set sequence as checked, so no StepID uniqueness is performed on next sequence execution
            _sut_N.SetSequenceAsChecked(); //Set sequence as checked, so no StepID uniqueness is performed on next sequence execution
            _sut_A.SetNumberOfSteps(10); //Set numberOfSteps to the testing instance
            _sut_N.SetNumberOfSteps(10); //Set numberOfSteps to the testing instance
            _sut_A.TcoSequencerTest := eTcoSequencerTests.RequestStep;
            _sut_N.TcoSequencerTest := eTcoSequencerTests.RequestStep;
            _plcCycleCounter := 0;
            _arranged := TRUE;
            RETURN;
        END_IF

        IF NOT _done THEN
            _sut_A.SequenceRun := _plcCycleCounter;
            _sut_N.SequenceRun := _plcCycleCounter;
            _sut_A.Run();
            _sut_N.Run();
        END_IF

        _done := _plcCycleCounter >= 3;
        ProbeDoneWhen(_done);
    {endregion}
    {region "T510_CheckStepIdUniqueness"}
    eTcoSequencerTests.CheckStepIdUniqueness:
        IF NOT _arranged THEN
            _sut_A.SetCyclicMode(); //Set sequencer into the cyclic mode
            _sut_N.SetCyclicMode(); //Set sequencer into the cyclic mode
            _sut_A.SetSequenceAsNotChecked(); //Set sequence as not checked, so StepId uniqueness is going to be performed on next sequence run
            _sut_N.SetSequenceAsNotChecked(); //Set sequence as not checked, so StepId uniqueness is going to be performed on next sequence run
            _sut_A.ClearNumberOfSteps(); //Clear internal step counters, so number of steps is going to be counted again on next sequence run
            _sut_N.ClearNumberOfSteps(); //Clear internal step counters, so number of steps is going to be counted again on next sequence run
            _sut_A.Enabled := TRUE;
            _sut_A.RunOneStep := FALSE;
            _sut_A.RunAllSteps := TRUE;
            _sut_A.FinishStep := TRUE;
            _sut_N.Enabled := TRUE;
            _sut_N.RunOneStep := FALSE;
            _sut_N.RunAllSteps := TRUE;
            _sut_N.FinishStep := TRUE;
            _sut_A.SetCurrentStep(inStepID := _currentStepId, inStepDescription := _currentStepDescription);
            _sut_N.SetCurrentStep(inStepID := _currentStepId, inStepDescription := _currentStepDescription);
            _sut_A.TcoSequencerTest := eTcoSequencerTests.CheckStepIdUniqueness;
            _sut_N.TcoSequencerTest := eTcoSequencerTests.CheckStepIdUniqueness;
            _sut_A.SaveNumberOfStepsInSequence();
            _sut_N.SaveNumberOfStepsInSequence();
            _plcCycleCounter := 0;
            _arranged := TRUE;
            RETURN;
        END_IF

        IF NOT _done THEN
            _sut_A.Run();
            _sut_N.Run();
            _sut_A.SaveNumberOfStepsInSequence();
            _sut_N.SaveNumberOfStepsInSequence();
        END_IF

        _done := _plcCycleCounter >= 2;
        ProbeDoneWhen(_done);
    {endregion}
    {region "T512_RestoreAlreadyCheckedSequence"}
    eTcoSequencerTests.RestoreAlreadyCheckedSequence:
        _sut_A.Restore();
        _sut_N.Restore();
        _sut_A.SaveNumberOfStepsInSequence();
        _sut_N.SaveNumberOfStepsInSequence();
        _done := TRUE;
        ProbeDoneWhen(_done);
    {endregion}
    {region "T513_CheckStepIdUniqueness"}
    eTcoSequencerTests.NotUniqueStepId:
        IF NOT _arranged THEN
            _sut_A.Enabled := TRUE;
            _sut_A.RunOneStep := FALSE;
            _sut_A.RunAllSteps := FALSE;
            _sut_A.FinishStep := TRUE;
            _sut_A.StepId := _stepId;
            _sut_N.Enabled := TRUE;
            _sut_N.RunOneStep := FALSE;
            _sut_N.RunAllSteps := FALSE;
            _sut_N.FinishStep := TRUE;
            _sut_N.StepId := _stepId;
            _sut_A.SetCurrentStep(inStepID := _currentStepId, inStepDescription := _currentStepDescription);
            _sut_N.SetCurrentStep(inStepID := _currentStepId, inStepDescription := _currentStepDescription);
            _sut_A.TcoSequencerTest := eTcoSequencerTests.NotUniqueStepId;
            _sut_N.TcoSequencerTest := eTcoSequencerTests.NotUniqueStepId;
            _sut_A.SaveNumberOfStepsInSequence();
            _sut_N.SaveNumberOfStepsInSequence();
            _plcCycleCounter := 0;
            _arranged := TRUE;
            RETURN;
        END_IF

        IF NOT _done THEN
            _sut_A.Run();
            _sut_N.Run();
            _sut_A.SaveNumberOfStepsInSequence();
            _sut_N.SaveNumberOfStepsInSequence();
            _done := _plcCycleCounter >= 2;
        END_IF

        IF _done THEN
            ProbeDoneWhen(_done);
        END_IF
    {endregion}
    {region "T516_AfterErrorRestore"}
    eTcoSequencerTests.AfterErrorRestore:
        IF NOT _arranged THEN
            _sut_A.TcoSequencerTest := eTcoSequencerTests.AfterErrorRestore;
            _sut_N.TcoSequencerTest := eTcoSequencerTests.AfterErrorRestore;
            _sut_A.SaveNumberOfStepsInSequence();
            _sut_N.SaveNumberOfStepsInSequence();
            _plcCycleCounter := 0;
            _arranged := TRUE;
            RETURN;
        END_IF

        IF NOT _done THEN
            _sut_A.Run();
            _sut_N.Run();
            _sut_A.SaveNumberOfStepsInSequence();
            _sut_N.SaveNumberOfStepsInSequence();
            _done := _plcCycleCounter >= 3;
        END_IF

        IF _done THEN
            ProbeDoneWhen(_done);
        END_IF
    {endregion}
    {region "T520_ChangeStepIdDuringExecution"}
    eTcoSequencerTests.ChangeStepIdDuringExecution:
        IF NOT _arranged THEN
            _sut_A.TcoSequencerTest := eTcoSequencerTests.ChangeStepIdDuringExecution;
            _sut_N.TcoSequencerTest := eTcoSequencerTests.ChangeStepIdDuringExecution;
            _sut_A.SetCyclicMode(); //Set sequencer into the cyclic mode
            _sut_N.SetCyclicMode(); //Set sequencer into the cyclic mode
            _sut_A.SetSequenceAsChecked(); //Set sequence as checked, so no StepID uniqueness is performed on next sequence execution
            _sut_N.SetSequenceAsChecked(); //Set sequence as checked, so no StepID uniqueness is performed on next sequence execution
            _sut_A.ClearNumberOfSteps(); //Clear internal step counters, so number of steps is going to be counted again on next sequence run
            _sut_N.ClearNumberOfSteps(); //Clear internal step counters, so number of steps is going to be counted again on next sequence run
            _sut_A.SetCurrentStep(inStepID := _currentStepId, inStepDescription := _currentStepDescription);
            _sut_N.SetCurrentStep(inStepID := _currentStepId, inStepDescription := _currentStepDescription);
            _sut_A.TotalStepNumber := _totalStepNumber;
            _sut_N.TotalStepNumber := _totalStepNumber;
            _sut_A.SaveNumberOfStepsInSequence();
            _sut_N.SaveNumberOfStepsInSequence();
            _plcCycleCounter := 0;
            _arranged := TRUE;
            RETURN;
        END_IF

        IF NOT _done THEN
            _sut_A.SequenceRun := _plcCycleCounter;
            _sut_N.SequenceRun := _plcCycleCounter;
            _sut_A.Run();
            _sut_N.Run();
            _sut_A.SaveNumberOfStepsInSequence();
            _sut_N.SaveNumberOfStepsInSequence();
        END_IF

        _done := _plcCycleCounter >= 3;
        ProbeDoneWhen(_done);
    {endregion}
    {region "T524_CommentOutPartOfRunningSequencer"}
    eTcoSequencerTests.CommentOutPartOfRunningSequencer:
        IF NOT _arranged THEN
            _sut_A.TcoSequencerTest := eTcoSequencerTests.CommentOutPartOfRunningSequencer;
            _sut_N.TcoSequencerTest := eTcoSequencerTests.CommentOutPartOfRunningSequencer;
            _sut_A.SetCyclicMode(); //Set sequencer into the cyclic mode
            _sut_N.SetCyclicMode(); //Set sequencer into the cyclic mode
            _sut_A.SetSequenceAsChecked(); //Set sequence as checked, so no StepID uniqueness is performed on next sequence execution
            _sut_N.SetSequenceAsChecked(); //Set sequence as checked, so no StepID uniqueness is performed on next sequence execution
            _sut_A.ClearNumberOfSteps(); //Clear internal step counters, so number of steps is going to be counted again on next sequence run
            _sut_N.ClearNumberOfSteps(); //Clear internal step counters, so number of steps is going to be counted again on next sequence run
            _sut_A.SetCurrentStep(inStepID := _currentStepId, inStepDescription := _currentStepDescription);
            _sut_N.SetCurrentStep(inStepID := _currentStepId, inStepDescription := _currentStepDescription);
            _sut_A.TotalStepNumber := _totalStepNumber;
            _sut_N.TotalStepNumber := _totalStepNumber;
            _sut_A.SaveNumberOfStepsInSequence();
            _sut_N.SaveNumberOfStepsInSequence();
            _plcCycleCounter := 0;
            _arranged := TRUE;
            RETURN;
        END_IF

        IF NOT _done THEN
            IF _plcCycleCounter = 3 THEN
                _sut_A.Restore();
                _sut_N.Restore();
                _sut_A.SetSequenceAsChecked(); //Set sequence as checked, so no StepID uniqueness is performed on next sequence execution
                _sut_N.SetSequenceAsChecked(); //Set sequence as checked, so no StepID uniqueness is performed on next sequence execution
                _sut_A.ClearNumberOfSteps(); //Clear internal step counters, so number of steps is going to be counted again on next sequence run
                _sut_N.ClearNumberOfSteps(); //Clear internal step counters, so number of steps is going to be counted again on next sequence run
            END_IF

            _sut_A.SequenceRun := _plcCycleCounter;
            _sut_N.SequenceRun := _plcCycleCounter;
            _sut_A.Run();
            _sut_N.Run();
            _sut_A.SaveNumberOfStepsInSequence();
            _sut_N.SaveNumberOfStepsInSequence();
        END_IF

        _done := _plcCycleCounter >= 3;
        ProbeDoneWhen(_done);
    {endregion}
    {region "T526_UncommentPartOfRunningSequencer"}
    eTcoSequencerTests.UncommentPartOfRunningSequencer:
        IF NOT _arranged THEN
            _sut_A.TcoSequencerTest := eTcoSequencerTests.UncommentPartOfRunningSequencer;
            _sut_N.TcoSequencerTest := eTcoSequencerTests.UncommentPartOfRunningSequencer;
            _sut_A.SetCyclicMode(); //Set sequencer into the cyclic mode
            _sut_N.SetCyclicMode(); //Set sequencer into the cyclic mode
            _sut_A.SetSequenceAsChecked(); //Set sequence as checked, so no StepID uniqueness is performed on next sequence execution
            _sut_N.SetSequenceAsChecked(); //Set sequence as checked, so no StepID uniqueness is performed on next sequence execution
            _sut_A.ClearNumberOfSteps(); //Clear internal step counters, so number of steps is going to be counted again on next sequence run
            _sut_N.ClearNumberOfSteps(); //Clear internal step counters, so number of steps is going to be counted again on next sequence run
            _sut_A.SetCurrentStep(inStepID := _currentStepId, inStepDescription := _currentStepDescription);
            _sut_N.SetCurrentStep(inStepID := _currentStepId, inStepDescription := _currentStepDescription);
            _sut_A.TotalStepNumber := _totalStepNumber;
            _sut_N.TotalStepNumber := _totalStepNumber;
            _sut_A.SaveNumberOfStepsInSequence();
            _sut_N.SaveNumberOfStepsInSequence();
            _plcCycleCounter := 0;
            _arranged := TRUE;
            RETURN;
        END_IF

        IF NOT _done THEN
            _sut_A.SequenceRun := _plcCycleCounter;
            _sut_N.SequenceRun := _plcCycleCounter;
            _sut_A.Run();
            _sut_N.Run();
            _sut_A.SaveNumberOfStepsInSequence();
            _sut_N.SaveNumberOfStepsInSequence();
        END_IF

        _done := _plcCycleCounter >= 2;
        ProbeDoneWhen(_done);
    {endregion}
    {region "T530_OpenCloseSequence"}
    eTcoSequencerTests.OpenCloseSequence:
        IF NOT _arranged THEN
            _sut_A.TcoSequencerTest := eTcoSequencerTests.OpenCloseSequence;
            _sut_N.TcoSequencerTest := eTcoSequencerTests.OpenCloseSequence;
            _sut_A.SetCyclicMode(); //Set sequencer into the cyclic mode
            _sut_N.SetCyclicMode(); //Set sequencer into the cyclic mode
            _sut_A.SetSequenceAsChecked(); //Set sequence as checked, so no StepID uniqueness is performed on next sequence execution
            _sut_N.SetSequenceAsChecked(); //Set sequence as checked, so no StepID uniqueness is performed on next sequence execution
            _sut_A.ClearNumberOfSteps(); //Clear internal step counters, so number of steps is going to be counted again on next sequence run
            _sut_N.ClearNumberOfSteps(); //Clear internal step counters, so number of steps is going to be counted again on next sequence run
            _sut_A.TotalStepNumber := _totalStepNumber;
            _sut_N.TotalStepNumber := _totalStepNumber;
            _sut_A.SaveNumberOfStepsInSequence();
            _sut_N.SaveNumberOfStepsInSequence();
            _plcCycleCounter := 0;
            _arranged := TRUE;
            RETURN;
        END_IF

        IF NOT _done THEN
            IF _plcCycleCounter = 1 THEN
                _sut_A.SequencerOpen();
                _sut_N.SequencerOpen();

                IF _sut_A._Step(0, TRUE, 'Step 0') THEN
                    _sut_A._StepCompleteWhen(TRUE);
                END_IF

                IF _sut_N._Step(0, TRUE, 'Step 0') THEN
                    _sut_N._StepCompleteWhen(TRUE);
                END_IF
            END_IF

            IF _plcCycleCounter = 2 THEN
                FOR i := 1 TO _totalStepNumber DO
                    _sut_A._Step(i, TRUE, CONCAT('Step ', INT_TO_STRING(i)));
                    _sut_N._Step(i, TRUE, CONCAT('Step ', INT_TO_STRING(i)));
                END_FOR

                _sut_A.SequencerClose();
                _sut_N.SequencerClose();
            END_IF

            IF _plcCycleCounter = 3 THEN
                _sut_A.SequencerOpen();
                _sut_N.SequencerOpen();
            END_IF

            IF _plcCycleCounter = 4 THEN
                IF _sut_A._Step(0, TRUE, 'Step 0') THEN
                    _sut_A._StepCompleteWhen(TRUE);
                END_IF

                IF _sut_N._Step(0, TRUE, 'Step 0') THEN
                    _sut_N._StepCompleteWhen(TRUE);
                END_IF
            END_IF

            IF _plcCycleCounter = 5 THEN
                FOR i := 1 TO _totalStepNumber DO
                    IF _sut_A._Step(i, TRUE, CONCAT('Step ', INT_TO_STRING(i))) THEN
                        _sut_A._StepCompleteWhen(TRUE);
                    END_IF

                    IF _sut_N._Step(i, TRUE, CONCAT('Step ', INT_TO_STRING(i))) THEN
                        _sut_N._StepCompleteWhen(TRUE);
                    END_IF
                END_FOR
            END_IF

            IF _plcCycleCounter = 6 THEN
                _sut_A._SequenceComplete();
                _sut_N._SequenceComplete();
                _sut_A.SequencerClose();
                _sut_N.SequencerClose();
            END_IF

            IF _plcCycleCounter = 7 THEN
                _sut_A.SequencerOpen();
                _sut_N.SequencerOpen();
            END_IF

            IF _plcCycleCounter = 8 THEN
                _sut_A.SequencerClose();
                _sut_N.SequencerClose();
            END_IF

            IF _plcCycleCounter = 9 THEN
                _sut_A.SequencerOpen();
                _sut_N.SequencerOpen();
                _sut_A._Step(0, TRUE, 'Step 0');
                _sut_N._Step(0, TRUE, 'Step 0');
                _sut_A.SequencerClose();
                _sut_N.SequencerClose();
            END_IF
        END_IF

        _done := _plcCycleCounter >= 9;
        ProbeDoneWhen(_done);
    {endregion}
    {region "T541_RequestStepFromLowerToHigher"}
    eTcoSequencerTests.RequestStepFromLowerToHigher:
        IF NOT _arranged THEN
            _sut_A.TcoSequencerTest := eTcoSequencerTests.RequestStepFromLowerToHigher;
            _sut_N.TcoSequencerTest := eTcoSequencerTests.RequestStepFromLowerToHigher;
            _sut_A.SetCyclicMode(); //Set sequencer into the cyclic mode
            _sut_N.SetCyclicMode(); //Set sequencer into the cyclic mode
            _sut_A.SetSequenceAsChecked(); //Set sequence as checked, so no StepID uniqueness is performed on next sequence execution
            _sut_N.SetSequenceAsChecked(); //Set sequence as checked, so no StepID uniqueness is performed on next sequence execution
            _sut_A.ClearNumberOfSteps(); //Clear internal step counters, so number of steps is going to be counted again on next sequence run
            _sut_N.ClearNumberOfSteps(); //Clear internal step counters, so number of steps is going to be counted again on next sequence run
            _sut_A.SetCurrentStep(inStepID := _currentStepId, inStepDescription := _currentStepDescription);
            _sut_N.SetCurrentStep(inStepID := _currentStepId, inStepDescription := _currentStepDescription);
            _sut_A.TotalStepNumber := _totalStepNumber;
            _sut_N.TotalStepNumber := _totalStepNumber;
            _sut_A.ReqStep := _reqStep;
            _sut_N.ReqStep := _reqStep;
            _sut_A.ReqStepNotExists := _reqStepNotExists;
            _sut_N.ReqStepNotExists := _reqStepNotExists;
            _sut_A.SaveNumberOfStepsInSequence();
            _sut_N.SaveNumberOfStepsInSequence();
            _plcCycleCounter := 0;
            _arranged := TRUE;
            RETURN;
        END_IF

        IF NOT _done THEN
            _sut_A.SequenceRun := _plcCycleCounter;
            _sut_N.SequenceRun := _plcCycleCounter;
            _sut_A.Run();
            _sut_N.Run();
            _sut_A.SaveNumberOfStepsInSequence();
            _sut_N.SaveNumberOfStepsInSequence();
        END_IF

        _done := _plcCycleCounter >= 2;
        ProbeDoneWhen(_done);
    {endregion}
    {region "T542_RequestStepFromHigherToLower"}
    eTcoSequencerTests.RequestStepFromHigherToLower:
        IF NOT _arranged THEN
            _sut_A.TcoSequencerTest := eTcoSequencerTests.RequestStepFromHigherToLower;
            _sut_N.TcoSequencerTest := eTcoSequencerTests.RequestStepFromHigherToLower;
            _sut_A.SetCyclicMode(); //Set sequencer into the cyclic mode
            _sut_N.SetCyclicMode(); //Set sequencer into the cyclic mode
            _sut_A.SetSequenceAsChecked(); //Set sequence as checked, so no StepID uniqueness is performed on next sequence execution
            _sut_N.SetSequenceAsChecked(); //Set sequence as checked, so no StepID uniqueness is performed on next sequence execution
            _sut_A.SetNumberOfSteps(_totalStepNumber);
            _sut_N.SetNumberOfSteps(_totalStepNumber);
            _sut_A.SetCurrentStep(inStepID := _currentStepId, inStepDescription := _currentStepDescription);
            _sut_N.SetCurrentStep(inStepID := _currentStepId, inStepDescription := _currentStepDescription);
            _sut_A.TotalStepNumber := _totalStepNumber;
            _sut_N.TotalStepNumber := _totalStepNumber;
            _sut_A.ReqStep := _reqStep;
            _sut_N.ReqStep := _reqStep;
            _sut_A.ReqStepNotExists := _reqStepNotExists;
            _sut_N.ReqStepNotExists := _reqStepNotExists;
            _sut_A.SaveNumberOfStepsInSequence();
            _sut_N.SaveNumberOfStepsInSequence();
            _plcCycleCounter := 0;
            _arranged := TRUE;
            RETURN;
        END_IF

        IF NOT _done THEN
            _sut_A.SequenceRun := _plcCycleCounter;
            _sut_N.SequenceRun := _plcCycleCounter;
            _sut_A.Run();
            _sut_N.Run();
            _sut_A.SaveNumberOfStepsInSequence();
            _sut_N.SaveNumberOfStepsInSequence();
        END_IF

        _done := _plcCycleCounter >= 2;
        ProbeDoneWhen(_done);
    {endregion}
    {region "T544_RequestStepToNotExistingStep"}
    eTcoSequencerTests.RequestStepToNotExistingStep:
        IF NOT _arranged THEN
            _sut_A.TcoSequencerTest := eTcoSequencerTests.RequestStepToNotExistingStep;
            _sut_N.TcoSequencerTest := eTcoSequencerTests.RequestStepToNotExistingStep;
            _sut_A.SetCyclicMode(); //Set sequencer into the cyclic mode
            _sut_N.SetCyclicMode(); //Set sequencer into the cyclic mode
            _sut_A.SetSequenceAsChecked(); //Set sequence as checked, so no StepID uniqueness is performed on next sequence execution
            _sut_N.SetSequenceAsChecked(); //Set sequence as checked, so no StepID uniqueness is performed on next sequence execution
            _sut_A.SetNumberOfSteps(_totalStepNumber);
            _sut_N.SetNumberOfSteps(_totalStepNumber);
            _sut_A.SetCurrentStep(inStepID := _currentStepId, inStepDescription := _currentStepDescription);
            _sut_N.SetCurrentStep(inStepID := _currentStepId, inStepDescription := _currentStepDescription);
            _sut_A.TotalStepNumber := _totalStepNumber;
            _sut_N.TotalStepNumber := _totalStepNumber;
            _sut_A.ReqStep := _reqStep;
            _sut_N.ReqStep := _reqStep;
            _sut_A.ReqStepNotExists := _reqStepNotExists;
            _sut_N.ReqStepNotExists := _reqStepNotExists;
            _sut_A.SaveNumberOfStepsInSequence();
            _sut_N.SaveNumberOfStepsInSequence();
            _plcCycleCounter := 0;
            _arranged := TRUE;
            RETURN;
        END_IF

        IF _plcCycleCounter = 4 THEN
            _sut_A.Restore();
            _sut_N.Restore();
            _sut_A.SetCyclicMode(); //Set sequencer into the cyclic mode
            _sut_N.SetCyclicMode(); //Set sequencer into the cyclic mode
            _sut_A.SetSequenceAsChecked(); //Set sequence as checked, so no StepID uniqueness is performed on next sequence execution
            _sut_N.SetSequenceAsChecked(); //Set sequence as checked, so no StepID uniqueness is performed on next sequence execution
            _sut_A.SetNumberOfSteps(_totalStepNumber);
            _sut_N.SetNumberOfSteps(_totalStepNumber);
            _sut_A.SetCurrentStep(inStepID := _currentStepId, inStepDescription := _currentStepDescription);
            _sut_N.SetCurrentStep(inStepID := _currentStepId, inStepDescription := _currentStepDescription);
            _sut_A.TotalStepNumber := _totalStepNumber;
            _sut_N.TotalStepNumber := _totalStepNumber;
        END_IF

        IF NOT _done THEN
            _sut_A.SequenceRun := _plcCycleCounter;
            _sut_N.SequenceRun := _plcCycleCounter;
            _sut_A.Run();
            _sut_N.Run();
            _sut_A.SaveNumberOfStepsInSequence();
            _sut_N.SaveNumberOfStepsInSequence();
        END_IF

        _done := _plcCycleCounter >= 4;
        ProbeDoneWhen(_done);
    {endregion}
    {region "T547_RequestStepWhilePreviousRequestStepHasNotBeenYetProcessed"}
    eTcoSequencerTests.RequestStepWhilePreviousRequestStepHasNotBeenYetProcessed:
        IF NOT _arranged THEN
            _sut_A.TcoSequencerTest := eTcoSequencerTests.RequestStepWhilePreviousRequestStepHasNotBeenYetProcessed;
            _sut_N.TcoSequencerTest := eTcoSequencerTests.RequestStepWhilePreviousRequestStepHasNotBeenYetProcessed;
            _sut_A.SetCyclicMode(); //Set sequencer into the cyclic mode
            _sut_N.SetCyclicMode(); //Set sequencer into the cyclic mode
            _sut_A.SetSequenceAsChecked(); //Set sequence as checked, so no StepID uniqueness is performed on next sequence execution
            _sut_N.SetSequenceAsChecked(); //Set sequence as checked, so no StepID uniqueness is performed on next sequence execution
            _sut_A.SetNumberOfSteps(_totalStepNumber);
            _sut_N.SetNumberOfSteps(_totalStepNumber);
            _sut_A.SetCurrentStep(inStepID := _currentStepId, inStepDescription := _currentStepDescription);
            _sut_N.SetCurrentStep(inStepID := _currentStepId, inStepDescription := _currentStepDescription);
            _sut_A.TotalStepNumber := _totalStepNumber;
            _sut_N.TotalStepNumber := _totalStepNumber;
            _sut_A.ReqStep := _reqStep;
            _sut_N.ReqStep := _reqStep;
            _sut_A.ReqStepNotExists := _reqStepNotExists;
            _sut_N.ReqStepNotExists := _reqStepNotExists;
            _sut_A.SaveNumberOfStepsInSequence();
            _sut_N.SaveNumberOfStepsInSequence();
            _plcCycleCounter := 0;
            _arranged := TRUE;
            RETURN;
        END_IF

        IF NOT _done THEN
            _sut_A.SequenceRun := _plcCycleCounter;
            _sut_N.SequenceRun := _plcCycleCounter;
            _sut_A.Run();
            _sut_N.Run();
            _sut_A.SaveNumberOfStepsInSequence();
            _sut_N.SaveNumberOfStepsInSequence();
        END_IF

        _done := TRUE;
        ProbeDoneWhen(_done);
    {endregion}
    {region "T551_DisableStepEnabledAndActiveInPreviousPLCcycle"}
    eTcoSequencerTests.DisableStepEnabledAndActiveInPreviousPLCcycle:
        IF NOT _arranged THEN
            _sut_A.TcoSequencerTest := eTcoSequencerTests.DisableStepEnabledAndActiveInPreviousPLCcycle;
            _sut_N.TcoSequencerTest := eTcoSequencerTests.DisableStepEnabledAndActiveInPreviousPLCcycle;
            _sut_A.SetCyclicMode(); //Set sequencer into the cyclic mode
            _sut_N.SetCyclicMode(); //Set sequencer into the cyclic mode
            _sut_A.SetSequenceAsChecked(); //Set sequence as checked, so no StepID uniqueness is performed on next sequence execution
            _sut_N.SetSequenceAsChecked(); //Set sequence as checked, so no StepID uniqueness is performed on next sequence execution
            _sut_A.SetNumberOfSteps(_totalStepNumber);
            _sut_N.SetNumberOfSteps(_totalStepNumber);
            _sut_A.TotalStepNumber := _totalStepNumber;
            _sut_N.TotalStepNumber := _totalStepNumber;
            _sut_A.SaveNumberOfStepsInSequence();
            _sut_N.SaveNumberOfStepsInSequence();
            _plcCycleCounter := 0;
            _arranged := TRUE;
            RETURN;
        END_IF

        IF NOT _done THEN
            IF _plcCycleCounter = 1 THEN
                _sut_A.SequencerOpen();

                IF _sut_A._Step(0, TRUE, 'Step 0') THEN
                    _sut_A._StepCompleteWhen(TRUE);
                END_IF

                FOR i := 1 TO _totalStepNumber - 2 DO
                    _sut_A._Step(i, TRUE, CONCAT('Step ', INT_TO_STRING(i)));
                END_FOR

                IF _sut_A._Step(_totalStepNumber - 1, TRUE, CONCAT('Step ', INT_TO_STRING(_totalStepNumber - 1))) THEN
                    _sut_A._SequenceComplete();
                END_IF

                _sut_A.SequencerClose();
                _sut_N.SequencerOpen();

                IF _sut_N._Step(0, TRUE, 'Step 0') THEN
                    _sut_N._StepCompleteWhen(TRUE);
                END_IF

                FOR i := 1 TO _totalStepNumber - 2 DO
                    _sut_N._Step(i, TRUE, CONCAT('Step ', INT_TO_STRING(i)));
                END_FOR

                IF _sut_N._Step(_totalStepNumber - 1, TRUE, CONCAT('Step ', INT_TO_STRING(_totalStepNumber - 1))) THEN
                    _sut_N._SequenceComplete();
                END_IF

                _sut_N.SequencerClose();
            END_IF

            IF _plcCycleCounter = 2 THEN
                _sut_A.SequencerOpen();

                IF _sut_A._Step(0, TRUE, 'Step 0') THEN
                    _sut_A._StepCompleteWhen(TRUE);
                END_IF

                IF _sut_A._Step(1, FALSE, 'Step 0') THEN
                    _sut_A._StepCompleteWhen(FALSE);
                END_IF

                _sut_N.SequencerOpen();

                IF _sut_N._Step(0, TRUE, 'Step 0') THEN
                    _sut_N._StepCompleteWhen(TRUE);
                END_IF

                IF _sut_N._Step(1, FALSE, 'Step 0') THEN
                    _sut_N._StepCompleteWhen(FALSE);
                END_IF
            END_IF

            IF _plcCycleCounter = 3 THEN
                FOR i := 2 TO _totalStepNumber - 1 DO
                    _sut_A._Step(i, TRUE, CONCAT('Step ', INT_TO_STRING(i)));
                END_FOR

                IF _sut_A._Step(_totalStepNumber, TRUE, CONCAT('Step ', INT_TO_STRING(_totalStepNumber))) THEN
                    _sut_A._SequenceComplete();
                END_IF

                _sut_A.SequencerClose();

                FOR i := 2 TO _totalStepNumber - 1 DO
                    _sut_N._Step(i, TRUE, CONCAT('Step ', INT_TO_STRING(i)));
                END_FOR

                IF _sut_N._Step(_totalStepNumber, TRUE, CONCAT('Step ', INT_TO_STRING(_totalStepNumber))) THEN
                    _sut_N._SequenceComplete();
                END_IF

                _sut_N.SequencerClose();
            END_IF

            _sut_A.SaveNumberOfStepsInSequence();
            _sut_N.SaveNumberOfStepsInSequence();
        END_IF

        _done := _plcCycleCounter >= 3;
        ProbeDoneWhen(_done);
    {endregion}
    {region "T560_RequestStepCallingCyclically"}
    eTcoSequencerTests.RequestStepCallingCyclically:
        IF NOT _arranged THEN
            _sut_A.TcoSequencerTest := eTcoSequencerTests.RequestStepCallingCyclically;
            _sut_N.TcoSequencerTest := eTcoSequencerTests.RequestStepCallingCyclically;
            _sut_A.SetCyclicMode(); //Set sequencer into the cyclic mode
            _sut_N.SetCyclicMode(); //Set sequencer into the cyclic mode
            _sut_A.SetSequenceAsChecked(); //Set sequence as checked, so no StepID uniqueness is performed on next sequence execution
            _sut_N.SetSequenceAsChecked(); //Set sequence as checked, so no StepID uniqueness is performed on next sequence execution
            _sut_A.SetNumberOfSteps(_totalStepNumber);
            _sut_N.SetNumberOfSteps(_totalStepNumber);
            _sut_A.TotalStepNumber := _totalStepNumber;
            _sut_N.TotalStepNumber := _totalStepNumber;
            _sut_A.InitReqStepCycle := _initReqStepCycle;
            _sut_N.InitReqStepCycle := _initReqStepCycle;
            _sut_A.SaveNumberOfStepsInSequence();
            _sut_N.SaveNumberOfStepsInSequence();
            _plcCycleCounter := 0;
            _arranged := TRUE;
            RETURN;
        END_IF

        IF NOT _done THEN
            IF _plcCycleCounter = 1 THEN
                _sut_A.SequencerOpen();
                _sut_N.SequencerOpen();
            END_IF

            IF _plcCycleCounter = 2 THEN
                _sut_A.SequencerOpen();
                _sut_A._RequestStep(10);
                _sut_A.SequencerClose();
                _sut_A.SequencerOpen();
                _sut_N.SequencerOpen();
                _sut_N._RequestStep(10);
                _sut_N.SequencerClose();
                _sut_N.SequencerOpen();
            END_IF

            IF _plcCycleCounter = 3 THEN
                _sut_A._Step(0, TRUE, 'Step 0');
                _sut_A._Step(20, TRUE, 'Step 20');
                _sut_A._Step(10, TRUE, 'Step 10');
                _sut_A.SequencerClose();
                _sut_N._Step(0, TRUE, 'Step 0');
                _sut_N._Step(20, TRUE, 'Step 20');
                _sut_N._Step(10, TRUE, 'Step 10');
                _sut_N.SequencerClose();
            END_IF

            IF _plcCycleCounter = 4 THEN
                _sut_A.InitReqStepCycle := _initReqStepCycle;
                _sut_N.InitReqStepCycle := _initReqStepCycle;
            END_IF

            IF _plcCycleCounter >= 5 THEN
                _sut_A.SequencerOpen();
                _sut_A.PostOpenRequestStepCycle := _sut_A.RequestStepCycle;
                _sut_A._Step(0, TRUE, 'Step 0');

                IF (_sut_A._Step(20, TRUE, 'Step 20')) THEN
                    _sut_A._RequestStep(20);
                END_IF

                IF (_sut_A._Step(10, TRUE, 'Step 10')) THEN
                    _sut_A._RequestStep(20);
                END_IF

                _sut_A.PreCloseRequestStepCycle := _sut_A.RequestStepCycle;
                _sut_A.SequencerClose();
                _sut_N.SequencerOpen();
                _sut_N.PostOpenRequestStepCycle := _sut_N.RequestStepCycle;
                _sut_N._Step(0, TRUE, 'Step 0');

                IF (_sut_N._Step(20, TRUE, 'Step 20')) THEN
                    _sut_N._RequestStep(20);
                END_IF

                IF (_sut_N._Step(10, TRUE, 'Step 10')) THEN
                    _sut_N._RequestStep(20);
                END_IF

                _sut_N.PreCloseRequestStepCycle := _sut_N.RequestStepCycle;
                _sut_N.SequencerClose();
            END_IF
        END_IF

        _sut_A.SaveNumberOfStepsInSequence();
        _sut_N.SaveNumberOfStepsInSequence();
        _done := _plcCycleCounter >= _cycles + 4;
        ProbeDoneWhen(_done);
    {endregion}
    {region "T570_SetStepMode"}
    eTcoSequencerTests.SetStepMode:
        IF NOT _arranged THEN
            _sut_A.TcoSequencerTest := eTcoSequencerTests.SetStepMode;
            _sut_N.TcoSequencerTest := eTcoSequencerTests.SetStepMode;
            _sut_A.SetStepMode(); //Set sequencer into the step mode
            _sut_N.SetStepMode(); //Set sequencer into the step mode
            _sut_A.SetSequenceAsChecked(); //Set sequence as checked, so no StepID uniqueness is performed on next sequence execution
            _sut_N.SetSequenceAsChecked(); //Set sequence as checked, so no StepID uniqueness is performed on next sequence execution
            _sut_A.ClearNumberOfSteps();
            _sut_N.ClearNumberOfSteps();
            _sut_A.SetCurrentStep(inStepID := _currentStepId, inStepDescription := _currentStepDescription);
            _sut_N.SetCurrentStep(inStepID := _currentStepId, inStepDescription := _currentStepDescription);
            _sut_A.TotalStepNumber := _totalStepNumber;
            _sut_N.TotalStepNumber := _totalStepNumber;
            _sut_A.SaveNumberOfStepsInSequence();
            _sut_N.SaveNumberOfStepsInSequence();
            _plcCycleCounter := 0;
            _arranged := TRUE;
            RETURN;
        END_IF

        IF NOT _done THEN
            _sut_A.SequenceRun := _plcCycleCounter;
            _sut_N.SequenceRun := _plcCycleCounter;

            IF _plcCycleCounter = 1 THEN
                _sut_A.Run();
                _sut_N.Run();
            END_IF

            IF _plcCycleCounter = 2 THEN
                _sut_A.SequencerOpen();
                _sut_A._StepIn();

                IF _sut_A._Step(0, TRUE, 'Initial step') THEN
                    _sut_A._StepCompleteWhen(TRUE);
                END_IF

                _sut_N.SequencerOpen();
                _sut_N._StepIn();

                IF _sut_N._Step(0, TRUE, 'Initial step') THEN
                    _sut_N._StepCompleteWhen(TRUE);
                END_IF
            END_IF

            IF _plcCycleCounter = 3 THEN
                IF _sut_A._Step(1, TRUE, 'Step 1') THEN
                    _sut_A._StepCompleteWhen(TRUE);
                END_IF

                IF _sut_N._Step(1, TRUE, 'Step 1') THEN
                    _sut_N._StepCompleteWhen(TRUE);
                END_IF

                FOR i := 2 TO _totalStepNumber - 2 DO
                    _sut_A._Step(i, TRUE, CONCAT('Step ', INT_TO_STRING(i)));
                    _sut_N._Step(i, TRUE, CONCAT('Step ', INT_TO_STRING(i)));
                END_FOR

                IF _sut_A._Step(_totalStepNumber - 1, TRUE, CONCAT('Step ', INT_TO_STRING(_totalStepNumber - 1))) THEN
                    _sut_A._SequenceComplete();
                END_IF

                IF _sut_N._Step(_totalStepNumber - 1, TRUE, CONCAT('Step ', INT_TO_STRING(_totalStepNumber - 1))) THEN
                    _sut_N._SequenceComplete();
                END_IF
            END_IF

            IF _plcCycleCounter = 4 THEN
                _sut_A.Run();
                _sut_N.Run();
            END_IF

            _sut_A.SaveNumberOfStepsInSequence();
            _sut_N.SaveNumberOfStepsInSequence();
        END_IF

        _done := _plcCycleCounter >= 4;
        ProbeDoneWhen(_done);
    {endregion}
    {region "T580_StepMode"}
    eTcoSequencerTests.StepMode:
        IF NOT _arranged THEN
            _sut_A.TcoSequencerTest := eTcoSequencerTests.StepMode;
            _sut_N.TcoSequencerTest := eTcoSequencerTests.StepMode;
            _sut_A.SetStepMode(); //Set sequencer into the step mode
            _sut_N.SetStepMode(); //Set sequencer into the step mode
            _sut_A.SetSequenceAsChecked(); //Set sequence as checked, so no StepID uniqueness is performed on next sequence execution
            _sut_N.SetSequenceAsChecked(); //Set sequence as checked, so no StepID uniqueness is performed on next sequence execution
            _sut_A.ClearNumberOfSteps();
            _sut_N.ClearNumberOfSteps();
            _sut_A.SetCurrentStep(inStepID := _currentStepId, inStepDescription := _currentStepDescription);
            _sut_N.SetCurrentStep(inStepID := _currentStepId, inStepDescription := _currentStepDescription);
            _sut_A.TotalStepNumber := _totalStepNumber;
            _sut_N.TotalStepNumber := _totalStepNumber;
            _sut_A.SaveNumberOfStepsInSequence();
            _sut_N.SaveNumberOfStepsInSequence();
            _plcCycleCounter := 0;
            _arranged := TRUE;
            RETURN;
        END_IF

        IF NOT _done THEN
            _sut_A.SequenceRun := _plcCycleCounter;
            _sut_N.SequenceRun := _plcCycleCounter;
            _sut_A.Run();
            _sut_N.Run();
            _sut_A.SaveNumberOfStepsInSequence();
            _sut_N.SaveNumberOfStepsInSequence();
        END_IF

        _done := _plcCycleCounter >= _totalStepNumber + 1;
        ProbeDoneWhen(_done);
    {endregion}
    {region "T582_InvalidMode"}
    eTcoSequencerTests.InvalidMode:
        IF NOT _arranged THEN
            _sut_A.TcoSequencerTest := eTcoSequencerTests.SetStepMode;
            _sut_N.TcoSequencerTest := eTcoSequencerTests.SetStepMode;
            _sut_A.SetCyclicMode(); //Set sequencer into the cyclic mode
            _sut_N.SetCyclicMode(); //Set sequencer into the cyclic mode
            _sut_A.SetSequenceAsChecked(); //Set sequence as checked, so no StepID uniqueness is performed on next sequence execution
            _sut_N.SetSequenceAsChecked(); //Set sequence as checked, so no StepID uniqueness is performed on next sequence execution
            _sut_A.SetNumberOfSteps(_totalStepNumber);
            _sut_N.SetNumberOfSteps(_totalStepNumber);
            _sut_A.SetCurrentStep(inStepID := _currentStepId, inStepDescription := _currentStepDescription);
            _sut_N.SetCurrentStep(inStepID := _currentStepId, inStepDescription := _currentStepDescription);
            _sut_A.TotalStepNumber := _totalStepNumber;
            _sut_N.TotalStepNumber := _totalStepNumber;
            _sut_A.SaveNumberOfStepsInSequence();
            _sut_N.SaveNumberOfStepsInSequence();
            _plcCycleCounter := 0;
            _arranged := TRUE;
            RETURN;
        END_IF

        IF NOT _done THEN
            _sut_A.SequenceRun := _plcCycleCounter;
            _sut_N.SequenceRun := _plcCycleCounter;

            IF _plcCycleCounter = 1 THEN
                _sut_A.SequencerOpen();
                _sut_N.SequencerOpen();

                FOR i := 0 TO _totalStepNumber - 1 DO
                    IF _sut_A._Step(i, TRUE, CONCAT('Step ', INT_TO_STRING(i))) THEN
                        _sut_A._StepCompleteWhen(TRUE);
                    END_IF

                    IF _sut_N._Step(i, TRUE, CONCAT('Step ', INT_TO_STRING(i))) THEN
                        _sut_N._StepCompleteWhen(TRUE);
                    END_IF
                END_FOR
            END_IF

            IF _plcCycleCounter = 2 THEN
                _sut_A._Step(_totalStepNumber, TRUE, CONCAT('Step ', INT_TO_STRING(_totalStepNumber)));
                _sut_N._Step(_totalStepNumber, TRUE, CONCAT('Step ', INT_TO_STRING(_totalStepNumber)));
                _sut_A.SequencerClose();
                _sut_N.SequencerClose();
            END_IF

            IF _plcCycleCounter = 3 THEN
                _sut_A.SequencerOpen();
                _sut_N.SequencerOpen();

                FOR i := 0 TO _totalStepNumber DO
                    _sut_A._Step(i, TRUE, CONCAT('Step ', INT_TO_STRING(i)));
                    _sut_N._Step(i, TRUE, CONCAT('Step ', INT_TO_STRING(i)));
                END_FOR

                _sut_A.SequencerClose();
                _sut_N.SequencerClose();
            END_IF

            _sut_A.SaveNumberOfStepsInSequence();
            _sut_N.SaveNumberOfStepsInSequence();
        END_IF

        _done := _plcCycleCounter >= 3;
        ProbeDoneWhen(_done);
    {endregion}
    {region "T582_StepInError"}
    eTcoSequencerTests.StepInError:
        IF NOT _arranged THEN
            _sut_A.TcoSequencerTest := eTcoSequencerTests.StepInError;
            _sut_N.TcoSequencerTest := eTcoSequencerTests.StepInError;
            _sut_A.SetCyclicMode(); //Set sequencer into the cyclic mode
            _sut_N.SetCyclicMode(); //Set sequencer into the cyclic mode
            _sut_A.SetSequenceAsChecked(); //Set sequence as checked, so no StepID uniqueness is performed on next sequence execution
            _sut_N.SetSequenceAsChecked(); //Set sequence as checked, so no StepID uniqueness is performed on next sequence execution
            _sut_A.SetNumberOfSteps(_totalStepNumber);
            _sut_N.SetNumberOfSteps(_totalStepNumber);
            _sut_A.SetCurrentStep(inStepID := _currentStepId, inStepDescription := _currentStepDescription);
            _sut_N.SetCurrentStep(inStepID := _currentStepId, inStepDescription := _currentStepDescription);
            _sut_A.TotalStepNumber := _totalStepNumber;
            _sut_N.TotalStepNumber := _totalStepNumber;
            _sut_A.SaveNumberOfStepsInSequence();
            _sut_N.SaveNumberOfStepsInSequence();
            _plcCycleCounter := 0;
            _arranged := TRUE;
            RETURN;
        END_IF

        IF NOT _done THEN
            _sut_A.SequenceRun := _plcCycleCounter;
            _sut_N.SequenceRun := _plcCycleCounter;

            IF _plcCycleCounter = 1 THEN
                _sut_A.SequencerOpen();
                _sut_N.SequencerOpen();

                FOR i := 0 TO _totalStepNumber - 1 DO
                    IF _sut_A._Step(i, TRUE, CONCAT('Step ', INT_TO_STRING(i))) THEN
                        _sut_A._StepCompleteWhen(TRUE);
                    END_IF

                    IF _sut_N._Step(i, TRUE, CONCAT('Step ', INT_TO_STRING(i))) THEN
                        _sut_N._StepCompleteWhen(TRUE);
                    END_IF
                END_FOR
            END_IF

            IF _plcCycleCounter = 2 THEN
                _sut_A._Step(_totalStepNumber, TRUE, CONCAT('Step ', INT_TO_STRING(_totalStepNumber)));
                _sut_N._Step(_totalStepNumber, TRUE, CONCAT('Step ', INT_TO_STRING(_totalStepNumber)));
                _sut_A.SequencerClose();
                _sut_N.SequencerClose();
            END_IF

            IF _plcCycleCounter = 3 THEN
                _sut_A.SequencerOpen();
                _sut_N.SequencerOpen();

                FOR i := 0 TO _totalStepNumber DO
                    _sut_A._Step(i, TRUE, CONCAT('Step ', INT_TO_STRING(i)));
                    _sut_N._Step(i, TRUE, CONCAT('Step ', INT_TO_STRING(i)));
                END_FOR

                _sut_A.SequencerClose();
                _sut_N.SequencerClose();
            END_IF

            _sut_A.SaveNumberOfStepsInSequence();
            _sut_N.SaveNumberOfStepsInSequence();
        END_IF

        _done := _plcCycleCounter >= 3;
        ProbeDoneWhen(_done);
    {endregion}
    {region "T590_CheckStepIdUniquenessStepMode"}
    eTcoSequencerTests.CheckStepIdUniquenessStepMode:
        IF NOT _arranged THEN
            _sut_A.SetStepMode(); //Set sequencer into the step mode
            _sut_N.SetStepMode(); //Set sequencer into the step mode
            _sut_A.SetSequenceAsNotChecked(); //Set sequence as not checked, so StepId uniqueness is going to be performed on next sequence run
            _sut_N.SetSequenceAsNotChecked(); //Set sequence as not checked, so StepId uniqueness is going to be performed on next sequence run
            _sut_A.ClearNumberOfSteps(); //Clear internal step counters, so number of steps is going to be counted again on next sequence run
            _sut_N.ClearNumberOfSteps(); //Clear internal step counters, so number of steps is going to be counted again on next sequence run
            _sut_A.Enabled := TRUE;
            _sut_A.RunOneStep := FALSE;
            _sut_A.RunAllSteps := TRUE;
            _sut_A.FinishStep := TRUE;
            _sut_A.StepId := _stepId;
            _sut_A.StepDescription := _stepDescription;
            _sut_N.Enabled := TRUE;
            _sut_N.RunOneStep := FALSE;
            _sut_N.RunAllSteps := TRUE;
            _sut_N.FinishStep := TRUE;
            _sut_N.StepId := _stepId;
            _sut_N.StepDescription := _stepDescription;
            _sut_A.SetCurrentStep(inStepID := _currentStepId, inStepDescription := _currentStepDescription);
            _sut_N.SetCurrentStep(inStepID := _currentStepId, inStepDescription := _currentStepDescription);
            _sut_A.TcoSequencerTest := eTcoSequencerTests.CheckStepIdUniquenessStepMode;
            _sut_N.TcoSequencerTest := eTcoSequencerTests.CheckStepIdUniquenessStepMode;
            _sut_A.SaveNumberOfStepsInSequence();
            _sut_N.SaveNumberOfStepsInSequence();
            _plcCycleCounter := 0;
            _arranged := TRUE;
            RETURN;
        END_IF

        IF NOT _done THEN
            IF _plcCycleCounter = 3 THEN
                _sut_A._StepIn();
                _sut_N._StepIn();
            END_IF

            _sut_A.Run();
            _sut_N.Run();

            IF _plcCycleCounter = 4 THEN
                _sut_A.Restore();
                _sut_N.Restore();
            END_IF

            _sut_A.SaveNumberOfStepsInSequence();
            _sut_N.SaveNumberOfStepsInSequence();
        END_IF

        _done := _plcCycleCounter >= 4;

        IF _done THEN
            _sut_A.TcoSequencerTest := eTcoSequencerTests.none;
            _sut_N.TcoSequencerTest := eTcoSequencerTests.none;
        END_IF

        ProbeDoneWhen(_done);
    {endregion}
    {region "T594_NotUniqueStepIdInStepMode"}
    eTcoSequencerTests.NotUniqueStepIdInStepMode:
        IF NOT _arranged THEN
            _sut_A.TcoSequencerTest := eTcoSequencerTests.NotUniqueStepIdInStepMode;
            _sut_N.TcoSequencerTest := eTcoSequencerTests.NotUniqueStepIdInStepMode;
            _sut_A.SetStepMode(); //Set sequencer into the step mode
            _sut_N.SetStepMode(); //Set sequencer into the step mode
            _sut_A.Enabled := TRUE;
            _sut_A.RunOneStep := FALSE;
            _sut_A.RunAllSteps := FALSE;
            _sut_A.FinishStep := TRUE;
            _sut_A.StepId := _stepId;
            _sut_N.Enabled := TRUE;
            _sut_N.RunOneStep := FALSE;
            _sut_N.RunAllSteps := FALSE;
            _sut_N.FinishStep := TRUE;
            _sut_N.StepId := _stepId;
            _sut_A.SetCurrentStep(inStepID := _currentStepId, inStepDescription := _currentStepDescription);
            _sut_N.SetCurrentStep(inStepID := _currentStepId, inStepDescription := _currentStepDescription);
            _sut_A.SaveNumberOfStepsInSequence();
            _sut_N.SaveNumberOfStepsInSequence();
            _plcCycleCounter := 0;
            _arranged := TRUE;
            RETURN;
        END_IF

        IF NOT _done THEN
            IF _plcCycleCounter = 2 THEN
                _Sut_A.RunOneStep := TRUE;
                _Sut_N.RunOneStep := TRUE;
            END_IF

            _sut_A.Run();
            _sut_N.Run();
            _sut_A.SaveNumberOfStepsInSequence();
            _sut_N.SaveNumberOfStepsInSequence();
            _done := _plcCycleCounter >= 2;
        END_IF

        IF _done THEN
            ProbeDoneWhen(_done);
        END_IF
    {endregion}
    {region "T597_AfterErrorResetInStepMode"}
    eTcoSequencerTests.AfterErrorResetInStepMode:
        IF NOT _arranged THEN
            _sut_A.TcoSequencerTest := eTcoSequencerTests.AfterErrorRestore;
            _sut_N.TcoSequencerTest := eTcoSequencerTests.AfterErrorRestore;
            _sut_A.SetStepMode();
            _sut_N.SetStepMode();
            _sut_A.SaveNumberOfStepsInSequence();
            _sut_N.SaveNumberOfStepsInSequence();
            _plcCycleCounter := 0;
            _arranged := TRUE;
            RETURN;
        END_IF

        IF NOT _done THEN
            IF _plcCycleCounter = 3 THEN
                _sut_A._StepIn();
                _sut_N._StepIn();
            END_IF

            _sut_A.Run();
            _sut_N.Run();
            _sut_A.SaveNumberOfStepsInSequence();
            _sut_N.SaveNumberOfStepsInSequence();
            _done := _plcCycleCounter >= 4;
        END_IF

        IF _done THEN
            ProbeDoneWhen(_done);
        END_IF
    {endregion}
    {region "T601_InvalidModeDetailed"}
    eTcoSequencerTests.InvalidModeDetailed:
        IF NOT _arranged THEN
            _sut_A.TcoSequencerTest := eTcoSequencerTests.InvalidModeDetailed;
            _sut_N.TcoSequencerTest := eTcoSequencerTests.InvalidModeDetailed;
            _sut_A.SetSequenceAsNotChecked();
            _sut_N.SetSequenceAsNotChecked();
            _sut_A.ClearNumberOfSteps();
            _sut_N.ClearNumberOfSteps();
            _sut_A.SetCurrentStep(_currentStepId, _currentStepDescription);
            _sut_N.SetCurrentStep(_currentStepId, _currentStepDescription);
            _sut_A.StepId := _stepId;
            _sut_N.StepId := _stepId;
            _sut_A.StepDescription := _stepDescription;
            _sut_N.StepDescription := _stepDescription;
            _sut_A.Enabled := TRUE;
            _sut_N.Enabled := TRUE;
            _sut_A.RunOneStep := FALSE;
            _sut_N.RunOneStep := FALSE;
            _sut_A.RunAllSteps := TRUE;
            _sut_N.RunAllSteps := TRUE;
            _sut_A.FinishStep := TRUE;
            _sut_N.FinishStep := TRUE;
            _sut_A.SetStepMode();
            _sut_N.SetStepMode();
            _sut_A.SaveNumberOfStepsInSequence();
            _sut_N.SaveNumberOfStepsInSequence();
            _plcCycleCounter := 0;
            _arranged := TRUE;
            RETURN;
        END_IF

        IF NOT _done THEN
            IF _plcCycleCounter = 2 THEN
                _sut_A.SetInvalidMode();
                _sut_N.SetInvalidMode();
                _sut_A.RunOneStep := TRUE;
                _sut_N.RunOneStep := TRUE;
                _sut_A.RunAllSteps := FALSE;
                _sut_N.RunAllSteps := FALSE;
            END_IF

            _sut_A.Run();
            _sut_N.Run();
            _sut_A.SaveNumberOfStepsInSequence();
            _sut_N.SaveNumberOfStepsInSequence();
            _done := _plcCycleCounter >= 2;
        END_IF

        IF _done THEN
            ProbeDoneWhen(_done);
        END_IF
    {endregion}
    {region "T604_StepInErrorDetailed"}
    eTcoSequencerTests.StepInErrorDetailed:
        IF NOT _arranged THEN
            _sut_A.TcoSequencerTest := eTcoSequencerTests.StepInErrorDetailed;
            _sut_N.TcoSequencerTest := eTcoSequencerTests.StepInErrorDetailed;
            _sut_A.SetSequenceAsNotChecked();
            _sut_N.SetSequenceAsNotChecked();
            _sut_A.ClearNumberOfSteps();
            _sut_N.ClearNumberOfSteps();
            _sut_A.SetCurrentStep(_currentStepId, _currentStepDescription);
            _sut_N.SetCurrentStep(_currentStepId, _currentStepDescription);
            _sut_A.StepId := _stepId;
            _sut_N.StepId := _stepId;
            _sut_A.StepDescription := _stepDescription;
            _sut_N.StepDescription := _stepDescription;
            _sut_A.Enabled := TRUE;
            _sut_N.Enabled := TRUE;
            _sut_A.RunOneStep := FALSE;
            _sut_N.RunOneStep := FALSE;
            _sut_A.RunAllSteps := TRUE;
            _sut_N.RunAllSteps := TRUE;
            _sut_A.FinishStep := TRUE;
            _sut_N.FinishStep := TRUE;
            _sut_A.SetStepMode();
            _sut_N.SetStepMode();
            _sut_A.SaveNumberOfStepsInSequence();
            _sut_N.SaveNumberOfStepsInSequence();
            _plcCycleCounter := 0;
            _arranged := TRUE;
            RETURN;
        END_IF

        IF NOT _done THEN
            IF _plcCycleCounter = 2 THEN
                _sut_A.SetCurrentStepToErrorState();
                _sut_N.SetCurrentStepToErrorState();
                _sut_A.RunOneStep := TRUE;
                _sut_N.RunOneStep := TRUE;
                _sut_A.RunAllSteps := FALSE;
                _sut_N.RunAllSteps := FALSE;
            END_IF

            _sut_A.Run();
            _sut_N.Run();
            _sut_A.SaveNumberOfStepsInSequence();
            _sut_N.SaveNumberOfStepsInSequence();
            _done := _plcCycleCounter >= 2;
        END_IF

        IF _done THEN
            ProbeDoneWhen(_done);
        END_IF
    {endregion}
    {region "T611_StepModeStepIn"}
    eTcoSequencerTests.StepModeStepIn:
        IF NOT _arranged THEN
            _sut_A.TcoSequencerTest := eTcoSequencerTests.StepModeStepIn;
            _sut_N.TcoSequencerTest := eTcoSequencerTests.StepModeStepIn;
            _sut_A.SetSequenceAsChecked();
            _sut_N.SetSequenceAsChecked();
            _sut_A.SetNumberOfSteps(_totalStepNumber);
            _sut_N.SetNumberOfSteps(_totalStepNumber);
            _sut_A.TotalStepNumber := _totalStepNumber;
            _sut_N.TotalStepNumber := _totalStepNumber;
            _sut_A.SetCurrentStep(_currentStepId, _currentStepDescription);
            _sut_N.SetCurrentStep(_currentStepId, _currentStepDescription);
            _sut_A.StepId := _stepId;
            _sut_N.StepId := _stepId;
            _sut_A.StepDescription := _stepDescription;
            _sut_N.StepDescription := _stepDescription;
            _sut_A.Enabled := TRUE;
            _sut_N.Enabled := TRUE;
            _sut_A.RunOneStep := FALSE;
            _sut_N.RunOneStep := FALSE;
            _sut_A.RunAllSteps := TRUE;
            _sut_N.RunAllSteps := TRUE;
            _sut_A.FinishStep := TRUE;
            _sut_N.FinishStep := TRUE;
            _sut_A.SetStepMode();
            _sut_N.SetStepMode();
            _sut_A.SaveNumberOfStepsInSequence();
            _sut_N.SaveNumberOfStepsInSequence();
            _plcCycleCounter := 0;
            _arranged := TRUE;
            RETURN;
        END_IF

        IF NOT _done THEN
            _sut_A.SequenceRun := _plcCycleCounter;
            _sut_N.SequenceRun := _plcCycleCounter;
            _sut_A.Run();
            _sut_N.Run();
            _sut_A.SaveNumberOfStepsInSequence();
            _sut_N.SaveNumberOfStepsInSequence();
            _done := _plcCycleCounter >= _totalStepNumber + 1;
        END_IF

        IF _done THEN
            ProbeDoneWhen(_done);
        END_IF
    {endregion}
    {region "T612_StepModeChangeStepIdDuringExecution"}
    eTcoSequencerTests.StepModeChangeStepIdDuringExecution:
        IF NOT _done AND _plcCycleCounter <= 2 THEN
            _sut_A.TcoSequencerTest := eTcoSequencerTests.StepModeChangeStepIdDuringExecution;
            _sut_N.TcoSequencerTest := eTcoSequencerTests.StepModeChangeStepIdDuringExecution;
            _sut_A.SequenceRun := _plcCycleCounter;
            _sut_N.SequenceRun := _plcCycleCounter;
            _sut_A.Run();
            _sut_N.Run();
            _sut_A.SaveNumberOfStepsInSequence();
            _sut_N.SaveNumberOfStepsInSequence();
        END_IF

        IF _plcCycleCounter >= 3 THEN
            _sut_A.Restore();
            _sut_N.Restore();
            _sut_A.SetSequenceAsChecked();
            _sut_N.SetSequenceAsChecked();
            _sut_A.SetNumberOfSteps(_totalStepNumber);
            _sut_N.SetNumberOfSteps(_totalStepNumber);
            _sut_A.TotalStepNumber := _totalStepNumber;
            _sut_N.TotalStepNumber := _totalStepNumber;
            _sut_A.SetStepMode();
            _sut_N.SetStepMode();
            _sut_A.SaveNumberOfStepsInSequence();
            _sut_N.SaveNumberOfStepsInSequence();
        END_IF

        _done := _plcCycleCounter >= 3;

        IF _done THEN
            ProbeDoneWhen(_done);
        END_IF
    {endregion}
    {region "T615_StepModeChangeStepOrder"}
    eTcoSequencerTests.StepModeChangeStepOrder:
        IF NOT _arranged THEN
            _sut_A.TcoSequencerTest := eTcoSequencerTests.StepModeChangeStepOrder;
            _sut_N.TcoSequencerTest := eTcoSequencerTests.StepModeChangeStepOrder;
            _sut_A.SetSequenceAsChecked();
            _sut_N.SetSequenceAsChecked();
            _sut_A.SetNumberOfSteps(_totalStepNumber);
            _sut_N.SetNumberOfSteps(_totalStepNumber);
            _sut_A.TotalStepNumber := _totalStepNumber;
            _sut_N.TotalStepNumber := _totalStepNumber;
            _sut_A.SetCurrentStep(_currentStepId, _currentStepDescription);
            _sut_N.SetCurrentStep(_currentStepId, _currentStepDescription);
            _sut_A.StepId := _stepId;
            _sut_N.StepId := _stepId;
            _sut_A.StepDescription := _stepDescription;
            _sut_N.StepDescription := _stepDescription;
            _sut_A.Enabled := TRUE;
            _sut_N.Enabled := TRUE;
            _sut_A.RunOneStep := FALSE;
            _sut_N.RunOneStep := FALSE;
            _sut_A.RunAllSteps := TRUE;
            _sut_N.RunAllSteps := TRUE;
            _sut_A.FinishStep := TRUE;
            _sut_N.FinishStep := TRUE;
            _sut_A.SetStepMode();
            _sut_N.SetStepMode();
            _sut_A.SaveNumberOfStepsInSequence();
            _sut_N.SaveNumberOfStepsInSequence();
            _plcCycleCounter := 0;
            _arranged := TRUE;
            RETURN;
        END_IF

        IF _plcCycleCounter <= _totalStepNumber + 2 THEN
            _sut_A.SequenceRun := _plcCycleCounter;
            _sut_N.SequenceRun := _plcCycleCounter;
            _sut_A.Run();
            _sut_N.Run();
            _sut_A.SaveNumberOfStepsInSequence();
            _sut_N.SaveNumberOfStepsInSequence();
        END_IF

        IF _plcCycleCounter >= _totalStepNumber + 3 THEN
            _sut_A.Restore();
            _sut_N.Restore();
            _sut_A.SetSequenceAsChecked();
            _sut_N.SetSequenceAsChecked();
            _sut_A.SetNumberOfSteps(_totalStepNumber);
            _sut_N.SetNumberOfSteps(_totalStepNumber);
            _sut_A.TotalStepNumber := _totalStepNumber;
            _sut_N.TotalStepNumber := _totalStepNumber;
            _sut_A.SetStepMode();
            _sut_N.SetStepMode();
            _sut_A.SaveNumberOfStepsInSequence();
            _sut_N.SaveNumberOfStepsInSequence();
        END_IF

        _done := _plcCycleCounter >= _totalStepNumber + 3;

